ACTION A_PassEmsCmd:
// MQTT 명령 받기 (EMS 지령원이 있는 현장): GVL_IF.g_stEmsCmd를 번호를 확인하며 복사해 지령원 FB_SrcEms에 넘김 (GVL_IF 머리말의 읽는 규칙)
// 번호가 홀수 = 쓰는 중, 복사 전후 번호가 다름 = 복사 중에 바뀜 → 이번 스캔은 지난 복사본 그대로 (다음 스캔에 다시 시도)
nEmsSeq := GVL_IF.g_nCmdSeq;
// [결함 10 되돌림 2026-11-04: 코드로 막지 않고 운영 규칙으로 해결 — EMS는 command 토픽을 retain=false로 발행 (retained 명령은 재구독 때 새 메시지로 와서 실행됨).
//   되돌린 수정: IF (nEmsSeq AND 1) = 0 AND nEmsSeq <> 0 THEN (번호 0을 유효로 보지 않음) → 재시작 뒤 처음 온 정상 명령까지 번호 맞추기에만 쓰여 버려지는 부작용이 있었음]
IF (nEmsSeq AND 1) = 0 THEN
	stEmsCopy := GVL_IF.g_stEmsCmd;
	IF GVL_IF.g_nCmdSeq = nEmsSeq THEN
		GVL_SITE.g_fbSrcEms.i_stCmd		:= stEmsCopy;
		GVL_SITE.g_fbSrcEms.i_bValid	:= TRUE;
	END_IF
END_IF
GVL_SITE.g_fbSrcEms.i_astUnitCfg	:= GVL_SITE.UNIT_CFG;
GVL_SITE.g_fbSrcEms.i_astBmsCfg		:= GVL_SITE.BMS_CFG;
// 스탠다드 스케줄 모드: EMS PCS 지령을 그 PCS의 유닛에 넘김 (한 PCS에 유닛이 여럿이면 정격 비율로 나눔). 모드는 유닛별 값을 냄
// [16번 수정 2026-11-09: 관리자가 접속점 그룹 단위가 되어 모드 하나(g_fbCmStdSched1)가 모든 유닛 칸을 받음. 원래 g_fbCmStdSched1 ← PCS1, g_fbCmStdSched2 ← PCS2 그대로]
// 살아 있음 = EMS 지령원 유효 (지난 스캔). P 지령은 FB_SrcEms.i_bPEnable(기본 FALSE)과 따로라, 둘을 같이 켜지 않음
stEmsOut := GVL_SITE.g_fbSrcEms.Output;
FOR nCmU := 1 TO GVL_PARAM.UNIT_COUNT DO
	nCmPcs := GVL_SITE.UNIT_CFG[nCmU].nPcs;
	IF nCmPcs >= 1 AND nCmPcs <= GVL_PARAM.PCS_COUNT THEN
		fCmPcsRated := 0.0;
		FOR nCmK := 1 TO GVL_PARAM.UNIT_COUNT DO
			IF GVL_SITE.UNIT_CFG[nCmK].nPcs = nCmPcs AND F_RealOk(GVL_SITE.UNIT_CFG[nCmK].fPRated) THEN
				fCmPcsRated := fCmPcsRated + MAX(GVL_SITE.UNIT_CFG[nCmK].fPRated, 0.0);
			END_IF
		END_FOR
		GVL_SITE.g_fbCmStdSched1.i_astCmd[nCmU].bUse		:= TRUE;
		GVL_SITE.g_fbCmStdSched1.i_astCmd[nCmU].bAlive		:= stEmsOut.bValid;
		GVL_SITE.g_fbCmStdSched1.i_astCmd[nCmU].nPSeq		:= stEmsCopy.anPcsPSeq[nCmPcs];
		IF fCmPcsRated > 0.0 AND F_RealOk(GVL_SITE.UNIT_CFG[nCmU].fPRated) THEN
			GVL_SITE.g_fbCmStdSched1.i_astCmd[nCmU].fP	:= stEmsCopy.afPcsP[nCmPcs] * MAX(GVL_SITE.UNIT_CFG[nCmU].fPRated, 0.0) / fCmPcsRated;
		ELSE
			GVL_SITE.g_fbCmStdSched1.i_astCmd[nCmU].fP	:= 0.0;
		END_IF
		GVL_SITE.g_fbCmStdSched1.i_astCmd[nCmU].nStateSeq	:= stEmsCopy.astPcs[nCmPcs].nSeq;
		GVL_SITE.g_fbCmStdSched1.i_astCmd[nCmU].eState		:= stEmsCopy.astPcs[nCmPcs].eCmd;
	ELSE
		GVL_SITE.g_fbCmStdSched1.i_astCmd[nCmU].bUse		:= FALSE;	// PCS 번호 범위 밖 (설정 점검 오류)
	END_IF
END_FOR
END_ACTION

ACTION A_Report:
// UPS site: no installed PCS. Do not publish a Plaspo mapping for a UPS.
GVL_IF.g_nReportSeq:=GVL_IF.g_nReportSeq+1;
FOR _nReportPcs:=1 TO GVL_PARAM.PCS_COUNT DO
 GVL_IF.g_stReport.abPcsMapped[_nReportPcs]:=FALSE;
 GVL_IF.g_stReport.abPcsComm[_nReportPcs]:=FALSE;
END_FOR
fbRptBat[1](i_stState:=GVL_SITE.g_fbBms1.q_stState, i_stRaw:=GVL_SITE.g_fbBms1.q_stRaw, i_nDeviceIndex:=1);	// BAT 번호 1부터 [1부터 2026-11-10]
FOR _nReportBat:=1 TO GVL_PARAM.BMS_COUNT DO
 GVL_IF.g_stReport.abBatMapped[_nReportBat]:=TRUE;
 GVL_IF.g_stReport.abBatValid[_nReportBat]:=fbRptBat[_nReportBat].q_bValid;
 GVL_IF.g_stReport.astBat[_nReportBat]:=fbRptBat[_nReportBat].q_stBat;
 FOR _nReportRack:=1 TO GVL_PARAM.RACKS_PER_BMS DO
  GVL_IF.g_stReport.astRack[(_nReportBat-1)*GVL_PARAM.RACKS_PER_BMS+_nReportRack]:=fbRptBat[_nReportBat].q_astRack[_nReportRack];
 END_FOR
 FOR _nReportModule:=1 TO GVL_PARAM.RACKS_PER_BMS*GVL_PARAM.MODULES_PER_RACK DO
  GVL_IF.g_stReport.astModule[(_nReportBat-1)*GVL_PARAM.RACKS_PER_BMS*GVL_PARAM.MODULES_PER_RACK+_nReportModule]:=fbRptBat[_nReportBat].q_astModule[_nReportModule];
 END_FOR
END_FOR
fbRptUps[1](i_stState:=GVL_SITE.g_fbUps1.q_stState, i_nDeviceIndex:=1);
FOR _nReportUps:=1 TO GVL_PARAM.UPS_COUNT DO
 GVL_IF.g_stReport.abUpsMapped[_nReportUps]:=TRUE;
 GVL_IF.g_stReport.abUpsValid[_nReportUps]:=fbRptUps[_nReportUps].q_bValid;
 GVL_IF.g_stReport.astUps[_nReportUps]:=fbRptUps[_nReportUps].q_stUps;
 // 명세 SQ-01: 사고·고장 단계. Fault 확인 = EMS UPS 명령 10 (WR-SQ-01)
 fbUpsSafety[_nReportUps](i_stUps:=fbRptUps[_nReportUps].q_stUps, i_bUpsValid:=fbRptUps[_nReportUps].q_bValid,
  i_stBat:=fbRptBat[_nReportUps].q_stBat, i_bBatValid:=fbRptBat[_nReportUps].q_bValid, i_bAck:=fbUpsCommand[_nReportUps].q_bAck);
END_FOR
// IMD 보고 (인터페이스 22. IMD)
fbRptImd[1](i_stState:=GVL_SITE.g_fbImd1.q_stState, i_nDeviceIndex:=1);
FOR _nReportImd:=1 TO GVL_PARAM.IMD_COUNT DO
 GVL_IF.g_stReport.abImdMapped[_nReportImd]:=TRUE;
 GVL_IF.g_stReport.abImdValid[_nReportImd]:=fbRptImd[_nReportImd].q_bValid;
 GVL_IF.g_stReport.astImd[_nReportImd]:=fbRptImd[_nReportImd].q_stImd;
END_FOR
// 화재감지기 보고 (토픽 fire_detector, 인터페이스 20. OffGas 양식: b0 통신 이상, b1 알람, b2 고장)
// 1 = TS-60 연기 접점 (g_fbIo1 DI 1, 통신 = EtherCAT 단자 상태), 2 = ASD-57 (연기 또는 온도 알람). 고장(b2)은 알 수 없어 0
GVL_IF.g_stReport.abFireMapped[1]:=TRUE;
GVL_IF.g_stReport.astFire[1].DeviceIndex:=1;
GVL_IF.g_stReport.astFire[1].Status:=SEL(GVL_SITE.g_fbIo1.Comm, UDINT#1, SEL(GVL_SITE.g_fbIo1.M_GetBit(i_nPoint:=1), UDINT#0, UDINT#2));
GVL_IF.g_stReport.abFireMapped[2]:=TRUE;
GVL_IF.g_stReport.astFire[2].DeviceIndex:=2;
GVL_IF.g_stReport.astFire[2].Status:=SEL(GVL_SITE.g_fbAsd57.q_bValid, UDINT#1, SEL(GVL_SITE.g_fbAsd57.q_bSmokeAlarm OR GVL_SITE.g_fbAsd57.q_bTempAlarm, UDINT#0, UDINT#2));
// 온습도 보고 (인터페이스 07.Temperature Sensor). location 2 = BAT실 (잠정, 현장 위치 확인)
fbRptTemp[1](i_stState:=GVL_SITE.g_fbThd2.q_stState, i_nDeviceIndex:=1, i_nLocation:=2);
GVL_IF.g_stReport.abTempMapped[1]:=TRUE;
GVL_IF.g_stReport.astTemp[1]:=fbRptTemp[1].q_stTemp;
GVL_IF.g_nReportSeq:=GVL_IF.g_nReportSeq+1;
END_ACTION

END_PROGRAM

// ---- 10_Core/10_Snapshot/FB_Snapshot.TcPOU
FUNCTION_BLOCK FB_Snapshot		// 이번 스캔의 장비 상태를 한 번에 복사. 이후 단계는 이 사본만 읽는다
VAR_IN_OUT
	iq_aipPcs		: ARRAY[1..GVL_PARAM.PCS_COUNT] OF I_Pcs;
	iq_aipBms		: ARRAY[1..GVL_PARAM.BMS_COUNT] OF I_Bms;
	iq_aipMeter		: ARRAY[1..GVL_PARAM.METER_COUNT] OF I_Meter;
END_VAR
VAR_IN_OUT CONSTANT
	iq_astUnitCfg	: ARRAY[1..GVL_PARAM.UNIT_COUNT] OF ST_UnitCfg;
END_VAR
VAR_OUTPUT
	q_astUnit		: ARRAY[1..GVL_PARAM.UNIT_COUNT] OF ST_UnitState;
	q_astBms		: ARRAY[1..GVL_PARAM.BMS_COUNT] OF ST_BatState;
	q_astMeter		: ARRAY[1..GVL_PARAM.METER_COUNT] OF ST_MeterState;
END_VAR
VAR_TEMP
	i				: UINT;
	nPcs			: UINT;
	stNoUnit		: ST_UnitState;		// 빈 칸: 통신 없음, 상태 Unknown
	stNoBms			: ST_BatState;
	stNoMeter		: ST_MeterState;
	k				: UINT;		// [결함 9 수정 2026-11-03: 추가]
END_VAR

// 유닛: 구성표의 PCS 번호·PCS 안 번호로 찾음
FOR i := 1 TO GVL_PARAM.UNIT_COUNT DO
	nPcs := iq_astUnitCfg[i].nPcs;
	IF nPcs >= 1 AND nPcs <= GVL_PARAM.PCS_COUNT AND_THEN iq_aipPcs[nPcs] <> 0 THEN
		q_astUnit[i] := iq_aipPcs[nPcs].M_GetUnitState(iq_astUnitCfg[i].nSub);
		q_astUnit[i].stP := M_FixVal(q_astUnit[i].stP);	// [결함 9 수정 2026-11-03: NaN·무한대 → 0·무효]
		q_astUnit[i].stQ := M_FixVal(q_astUnit[i].stQ);
	ELSE
		q_astUnit[i] := stNoUnit;
	END_IF
END_FOR

FOR i := 1 TO GVL_PARAM.BMS_COUNT DO
	IF iq_aipBms[i] <> 0 THEN
		q_astBms[i] := iq_aipBms[i].BatState;
		q_astBms[i].stSoc := M_FixVal(q_astBms[i].stSoc);	// [결함 9 수정 2026-11-03: NaN·무한대 → 0·무효, 한도는 0]
		q_astBms[i].stSoh := M_FixVal(q_astBms[i].stSoh);
		IF NOT F_CmdOk(q_astBms[i].fPChgMax, 0.0) THEN q_astBms[i].fPChgMax := 0.0; END_IF
		IF NOT F_CmdOk(q_astBms[i].fPDisMax, 0.0) THEN q_astBms[i].fPDisMax := 0.0; END_IF
	ELSE
		q_astBms[i] := stNoBms;
	END_IF
END_FOR

FOR i := 1 TO GVL_PARAM.METER_COUNT DO
	IF iq_aipMeter[i] <> 0 THEN
		q_astMeter[i] := iq_aipMeter[i].MeterState;
		q_astMeter[i].stP := M_FixVal(q_astMeter[i].stP);	// [결함 9 수정 2026-11-03: NaN·무한대 → 0·무효]
		q_astMeter[i].stQ := M_FixVal(q_astMeter[i].stQ);
		q_astMeter[i].stV := M_FixVal(q_astMeter[i].stV);
		FOR k := 1 TO 3 DO
			q_astMeter[i].astV[k] := M_FixVal(q_astMeter[i].astV[k]);
		END_FOR
		q_astMeter[i].stF := M_FixVal(q_astMeter[i].stF);
	ELSE
		q_astMeter[i] := stNoMeter;
	END_IF
END_FOR

METHOD PRIVATE M_FixVal : ST_Val		// 장비 값이 NaN·무한대면 0·무효로 (뒤 계산·비교에 퍼지지 않게). [결함 9 수정 2026-11-03: 추가]
VAR_INPUT
	i_stVal	: ST_Val;
END_VAR
M_FixVal := i_stVal;
IF NOT F_CmdOk(i_stVal.fValue, 0.0) THEN
	M_FixVal.fValue	:= 0.0;
	M_FixVal.bValid	:= FALSE;
END_IF
END_METHOD

END_FUNCTION_BLOCK

// ---- 10_Core/40_Arbitration/F_CmdOk.TcPOU
FUNCTION F_CmdOk : BOOL		// 지령값이 쓸 만한가: NaN·무한대가 아니고, 한도가 있으면 |값| ≤ 한도
VAR_INPUT
	i_fValue	: REAL;
	i_fLimit	: REAL;			// 0 이하 = 한도 검사 안 함
END_VAR

// NaN·무한대는 비트로 먼저 거름 (NaN을 크기 비교하면 PLC가 멈춤). 크기 비교는 보통 숫자일 때만
// [2026-11-05 머지: main의 F_IsFinite 방식 + 1.0E30 상한은 원래 코드대로 남김. 통합시험 결함 9 수정(비트 검사·dwBits)은 이 방식으로 합침]
F_CmdOk := F_IsFinite(i_fValue) AND_THEN ABS(i_fValue) < 1.0E30;
IF F_CmdOk AND i_fLimit > 0 THEN
	F_CmdOk := ABS(i_fValue) <= i_fLimit;
END_IF

END_FUNCTION

// ---- 10_Core/10_Snapshot/FB_Measure.TcPOU
FUNCTION_BLOCK FB_Measure		// 계측점 계산 + 제어 그룹마다 접속점 값·가상신호
VAR_INPUT
	i_bTestMode		: BOOL;			// 시험 모드에서만 가상신호를 씀 (GVL_SITE.TEST_MODE)
END_VAR
VAR_IN_OUT CONSTANT
	iq_astMeter		: ARRAY[1..GVL_PARAM.METER_COUNT] OF ST_MeterState;
	iq_astPointCfg	: ARRAY[1..GVL_PARAM.POINT_COUNT] OF ST_PointCfg;
	iq_astGroupCfg	: ARRAY[1..GVL_PARAM.GROUP_COUNT] OF ST_GroupCfg;
	iq_astVirtual	: ARRAY[1..GVL_PARAM.GROUP_COUNT] OF ST_VirtualSet;
END_VAR
VAR_OUTPUT
	q_astPoint		: ARRAY[1..GVL_PARAM.POINT_COUNT] OF ST_MeterState;	// 계측점 (실측, 가상신호 적용 전)
	q_astPcc		: ARRAY[1..GVL_PARAM.GROUP_COUNT] OF ST_PccMeas;		// 그룹 접속점 (가상신호 적용 후)
END_VAR
VAR_TEMP
	nPointNo				: UINT;
	nTermNo				: UINT;
	g				: UINT;
	k				: UINT;
	nMeterNo				: UINT;
	bFirst			: BOOL;		// 아직 묶인 계측기를 못 만남
	bComm			: BOOL;
	bPValid			: BOOL;
	bQValid			: BOOL;
	stPoint			: ST_MeterState;
	stNone			: ST_MeterState;	// 빈 값: 통신 없음, 값 무효
END_VAR

(* 1) 계측점: 계측기 P·Q를 부호와 함께 더함. 전압·주파수는 첫 계측기 값 *)
FOR nPointNo := 1 TO GVL_PARAM.POINT_COUNT DO
	stPoint	:= stNone;
	bFirst	:= TRUE;
	bComm	:= TRUE;
	bPValid	:= TRUE;
	bQValid	:= TRUE;
	FOR nTermNo := 1 TO GVL_PARAM.POINT_TERM_MAX DO
		nMeterNo := iq_astPointCfg[nPointNo].astTerm[nTermNo].nMeter;
		IF nMeterNo > GVL_PARAM.METER_COUNT THEN
			bComm := FALSE;		// 설정 오류: 없는 계측기
		ELSIF nMeterNo >= 1 THEN
			IF bFirst THEN
				stPoint.stV	:= iq_astMeter[nMeterNo].stV;
				stPoint.astV	:= iq_astMeter[nMeterNo].astV;
				stPoint.stF	:= iq_astMeter[nMeterNo].stF;
				bFirst		:= FALSE;
			END_IF
			bComm			:= bComm AND iq_astMeter[nMeterNo].bComm;
			bPValid			:= bPValid AND iq_astMeter[nMeterNo].stP.bValid;
			bQValid			:= bQValid AND iq_astMeter[nMeterNo].stQ.bValid;
			stPoint.stP.fValue	:= stPoint.stP.fValue + iq_astPointCfg[nPointNo].astTerm[nTermNo].fSign * iq_astMeter[nMeterNo].stP.fValue;
			stPoint.stQ.fValue	:= stPoint.stQ.fValue + iq_astPointCfg[nPointNo].astTerm[nTermNo].fSign * iq_astMeter[nMeterNo].stQ.fValue;
		END_IF
	END_FOR
	// 묶인 계측기가 없거나 하나라도 끊기면 무효
	stPoint.bComm		:= bComm AND NOT bFirst;
	stPoint.stP.bValid	:= stPoint.bComm AND bPValid;
	stPoint.stQ.bValid	:= stPoint.bComm AND bQValid;
	q_astPoint[nPointNo]	:= stPoint;
END_FOR

(* 2) 그룹 접속점 + 가상신호 *)
FOR g := 1 TO GVL_PARAM.GROUP_COUNT DO
	nPointNo := iq_astGroupCfg[g].nPccPoint;
	q_astPcc[g].bNoPoint := nPointNo = 0;	// [결함 7 수정 2026-11-03: 추가. 접속점 무효 보호가 '없음'을 무효로 보지 않게]
	IF nPointNo >= 1 AND nPointNo <= GVL_PARAM.POINT_COUNT THEN
		q_astPcc[g].stMeas := q_astPoint[nPointNo];
	ELSE
		q_astPcc[g].stMeas := stNone;
	END_IF

	// 가상 전압: 평균·상전압 모두 같은 값
	IF i_bTestMode AND iq_astVirtual[g].bVEna THEN
		q_astPcc[g].stMeas.stV.fValue	:= iq_astVirtual[g].fV;
		q_astPcc[g].stMeas.stV.bValid	:= TRUE;
		FOR k := 1 TO 3 DO
			q_astPcc[g].stMeas.astV[k].fValue	:= iq_astVirtual[g].fV;
			q_astPcc[g].stMeas.astV[k].bValid	:= TRUE;
		END_FOR
	END_IF

	// 가상 유효전력
	IF i_bTestMode AND iq_astVirtual[g].bPEna THEN
		q_astPcc[g].stMeas.stP.fValue	:= iq_astVirtual[g].fP;
		q_astPcc[g].stMeas.stP.bValid	:= TRUE;
	END_IF
END_FOR

END_FUNCTION_BLOCK

// ---- 10_Core/20_Protection/FB_Protection.TcPOU
FUNCTION_BLOCK FB_Protection		// 등록된 보호 칸마다 대상마다: 조건 모듈 판단 → 같은 칸 대응 모듈 → 유닛·BMS마다 요청 합치기 (센 조치·낮은 상한, 건 모듈 ID). 요청만, 장비에 직접 명령하지 않음
// 지연 없음: 통신 에러·고장은 장비 쪽(드라이버)이 판정해 올림. 현장 접점·아날로그의 떨림 방지는 조건 모듈 설정에
// 보호는 조건이 있는 동안만 걸림 (래치 없음). 다시 돌지 않아야 하면 정지나 Manual 전환을 씀
VAR_IN_OUT CONSTANT
	iq_astUnit		: ARRAY[1..GVL_PARAM.UNIT_COUNT] OF ST_UnitState;
	iq_astBms		: ARRAY[1..GVL_PARAM.BMS_COUNT] OF ST_BatState;
	iq_astPcc		: ARRAY[1..GVL_PARAM.GROUP_COUNT] OF ST_PccMeas;
	iq_astUnitCfg	: ARRAY[1..GVL_PARAM.UNIT_COUNT] OF ST_UnitCfg;
	iq_astBmsCfg	: ARRAY[1..GVL_PARAM.BMS_COUNT] OF ST_BmsCfg;
	iq_astRuleCfg	: ARRAY[1..GVL_PARAM.RULE_COUNT] OF ST_RuleCfg;
	iq_abUnitInstalled	: ARRAY[1..GVL_PARAM.UNIT_COUNT] OF BOOL;	// 미설치(칸 비어 있음)는 모듈에 bInstalled = FALSE로 넘김 (FB_ModuleList)
	iq_abBmsInstalled	: ARRAY[1..GVL_PARAM.BMS_COUNT] OF BOOL;
	iq_aeOpMode		: ARRAY[1..GVL_PARAM.UNIT_COUNT] OF E_OpMode;		// 실제 운전 모드 (대응이 그 모드 유닛에 조치를 걸지 봄)
END_VAR
VAR_IN_OUT
	iq_aipRule		: ARRAY[1..GVL_PARAM.RULE_COUNT] OF I_ProtectionRule;	// 조건 모듈
	iq_aipResp		: ARRAY[1..GVL_PARAM.RULE_COUNT] OF I_ProtResponse;	// 대응 모듈 (같은 칸). 비우면 조치 없음 (알람만)
END_VAR
VAR_OUTPUT
	q_astUnitProt	: ARRAY[1..GVL_PARAM.UNIT_COUNT] OF ST_UnitProt;		// 유닛별 가장 센 PCS 조치·가장 낮은 P·Q 상한·Manual 전환
	q_astBmsProt	: ARRAY[1..GVL_PARAM.BMS_COUNT] OF ST_BmsProt;		// BMS별 가장 센 배터리 조치
	q_aabRule		: ARRAY[1..GVL_PARAM.RULE_COUNT, 1..GVL_PARAM.PROT_TARGET_MAX] OF BOOL;	// 보호 발생 [규칙 칸, 대상 번호] (온라인 확인·로그용). Site는 대상 1
END_VAR
VAR
	_aatonActive	: ARRAY[1..GVL_PARAM.RULE_COUNT, 1..GVL_PARAM.PROT_TARGET_MAX] OF TON;	// 조건이 이어진 시간 (대응에 넘김)
	_stView			: ST_ProtView;		// 마지막으로 조건 모듈에 넘긴 정보 (온라인 확인용)
	_stReq			: ST_ProtReq;		// 마지막 대응 요청 (온라인 확인용)
	_stNoReq		: ST_ProtReq;		// 요청 없음 (비우기용. 처음 한 번 P·Q 상한을 100으로)
	_bInit			: BOOL;
END_VAR
VAR_TEMP
	i				: UINT;		// 규칙 칸
	t				: UINT;		// 대상 번호
	nTargetCount	: UINT;		// 이 규칙 범위의 대상 수
	bInRange		: BOOL;		// 이 대상을 보는가
	bCond			: BOOL;
	nModule			: UINT;
	stNoUnit		: ST_UnitProt;
	stNoBms			: ST_BmsProt;
	stNoView		: ST_ProtView;
END_VAR

(* 0) 이번 스캔 결과 비우기 *)
IF NOT _bInit THEN
	FOR i := 1 TO GVL_PARAM.UNIT_COUNT DO
		_stNoReq.afPPct[i] := 100.0;
		_stNoReq.afQPct[i] := 100.0;
	END_FOR
	_bInit := TRUE;
END_IF
FOR i := 1 TO GVL_PARAM.UNIT_COUNT DO
	q_astUnitProt[i] := stNoUnit;
END_FOR
FOR i := 1 TO GVL_PARAM.BMS_COUNT DO
	q_astBmsProt[i] := stNoBms;
END_FOR
(* 1) 보호 규칙 칸마다, 범위 안 대상마다: 조건 모듈 → 대응 → 합치기
   대상 번호(nTarget) 0 = 범위 안 대상 전부를 하나씩 (유닛 범위면 유닛 1..UNIT_COUNT). Site는 대상 1 하나 *)
FOR i := 1 TO GVL_PARAM.RULE_COUNT DO
	CASE iq_astRuleCfg[i].eScope OF
		E_ProtScope.Unit:		nTargetCount := GVL_PARAM.UNIT_COUNT;
		E_ProtScope.Bms:		nTargetCount := GVL_PARAM.BMS_COUNT;
		E_ProtScope.BatGroup:	nTargetCount := GVL_PARAM.BAT_COUNT;
		E_ProtScope.Group:		nTargetCount := GVL_PARAM.GROUP_COUNT;
	ELSE
		nTargetCount := 1;		// Site
	END_CASE
	nModule := 0;
	IF iq_aipRule[i] <> 0 THEN
		nModule := iq_aipRule[i].ModuleId;
	END_IF
	FOR t := 1 TO GVL_PARAM.PROT_TARGET_MAX DO
		bInRange := iq_aipRule[i] <> 0 AND t <= nTargetCount
			AND (iq_astRuleCfg[i].nTarget = 0 OR iq_astRuleCfg[i].nTarget = t OR iq_astRuleCfg[i].eScope = E_ProtScope.Site);
		bCond := FALSE;
		IF bInRange THEN
			// 조건 모듈에 넘길 정보: 범위·대상 번호·임계값과 그 대상의 상태
			_stView				:= stNoView;
			_stView.eScope		:= iq_astRuleCfg[i].eScope;
			_stView.nTarget		:= t;
			_stView.fThreshold	:= iq_astRuleCfg[i].fThreshold;
			_stView.bInstalled	:= TRUE;
			CASE iq_astRuleCfg[i].eScope OF
				E_ProtScope.Unit:
					_stView.bInstalled	:= iq_abUnitInstalled[t];
					_stView.stUnit		:= iq_astUnit[t];
					_stView.eOpMode		:= iq_aeOpMode[t];
					_stView.nGroup		:= iq_astUnitCfg[t].nGroup;
					_stView.nBatGroup	:= iq_astUnitCfg[t].nBatGroup;
				E_ProtScope.Bms:
					_stView.bInstalled	:= iq_abBmsInstalled[t];
					_stView.stBms		:= iq_astBms[t];
					_stView.nBatGroup	:= iq_astBmsCfg[t].nBatGroup;
				E_ProtScope.BatGroup:
					_stView.nBatGroup	:= t;
				E_ProtScope.Group:
					_stView.stPcc		:= iq_astPcc[t];
					_stView.nGroup		:= t;
			END_CASE
			// 등록 bAuto·bManual 중 하나라도 켜져 있어야 감지 (둘 다 끄면 이 보호를 안 씀)
			bCond := (iq_astRuleCfg[i].stProt.bAuto OR iq_astRuleCfg[i].stProt.bManual) AND iq_aipRule[i].M_Evaluate(_stView);
		END_IF
		q_aabRule[i, t] := bCond;
		_aatonActive[i, t](IN := bCond, PT := T#24D);
		// 대응: 매 스캔 부름 (조건이 없을 때도: 단계 대응이 풀린 뒤 상태를 정리할 수 있게). 대응 칸이 비면 조치 없음 (알람만)
		IF bInRange AND iq_aipResp[i] <> 0 THEN
			_stReq := _stNoReq;
			iq_aipResp[i].M_Respond(i_bActive := bCond, i_tActive := _aatonActive[i, t].ET, i_nTarget := t, i_stRule := iq_astRuleCfg[i],
				iq_astUnit := iq_astUnit, iq_astBms := iq_astBms, iq_astUnitCfg := iq_astUnitCfg, iq_astBmsCfg := iq_astBmsCfg,
				iq_aeOpMode := iq_aeOpMode, iq_stReq := _stReq);
			M_Merge(nModule);
		END_IF
	END_FOR
END_FOR

METHOD PRIVATE M_Merge		// 대응 요청(_stReq)을 장비마다 합침: PCS·배터리는 센 쪽, P·Q 상한은 낮은 쪽, Manual 전환은 하나라도. 건 모듈 = 조건 모듈 ID
VAR_INPUT
	i_nModule	: UINT;
END_VAR
VAR
	u			: UINT;
	m			: UINT;
END_VAR
FOR u := 1 TO GVL_PARAM.UNIT_COUNT DO
	IF F_PcsRank(_stReq.aePcs[u]) > F_PcsRank(q_astUnitProt[u].ePcsAction) THEN
		q_astUnitProt[u].ePcsAction	:= _stReq.aePcs[u];
		q_astUnitProt[u].nModule	:= i_nModule;
	END_IF
	IF _stReq.abToManual[u] AND NOT q_astUnitProt[u].bModeManualReq THEN
		q_astUnitProt[u].bModeManualReq	:= TRUE;
		q_astUnitProt[u].nModeModule	:= i_nModule;
	END_IF
	IF _stReq.afPPct[u] < q_astUnitProt[u].fPPct THEN
		q_astUnitProt[u].fPPct		:= _stReq.afPPct[u];
		q_astUnitProt[u].nPModule	:= i_nModule;
	END_IF
	IF _stReq.afQPct[u] < q_astUnitProt[u].fQPct THEN
		q_astUnitProt[u].fQPct		:= _stReq.afQPct[u];
		q_astUnitProt[u].nQModule	:= i_nModule;
	END_IF
END_FOR
FOR m := 1 TO GVL_PARAM.BMS_COUNT DO
	IF F_BatRank(_stReq.aeBat[m]) > F_BatRank(q_astBmsProt[m].eBatAction) THEN
		q_astBmsProt[m].eBatAction	:= _stReq.aeBat[m];
		q_astBmsProt[m].nModule		:= i_nModule;
	END_IF
END_FOR
END_METHOD

END_FUNCTION_BLOCK

// ---- 10_Core/20_Protection/F_PcsRank.TcPOU
FUNCTION F_PcsRank : INT		// 조치 세기: None 0 < Standby 1 < Stop 2 < EStop 3
VAR_INPUT
	i_eAction	: E_PcsAction;
END_VAR

CASE i_eAction OF
	E_PcsAction.Standby:	F_PcsRank := 1;
	E_PcsAction.Stop:		F_PcsRank := 2;
	E_PcsAction.EStop:		F_PcsRank := 3;
ELSE
	F_PcsRank := 0;
END_CASE

END_FUNCTION

// ---- 10_Core/20_Protection/F_BatRank.TcPOU
FUNCTION F_BatRank : INT		// 조치 세기: None 0 < Stop 1 < EStop 2
VAR_INPUT
	i_eAction	: E_BatAction;
END_VAR

CASE i_eAction OF
	E_BatAction.Stop:	F_BatRank := 1;
	E_BatAction.EStop:	F_BatRank := 2;
ELSE
	F_BatRank := 0;
END_CASE

END_FUNCTION

// ---- 10_Core/20_Protection/FB_BatGroup.TcPOU
FUNCTION_BLOCK FB_BatGroup		// BMS마다 쓸 수 있는지 판단, 배터리 그룹(DC 버스)마다 쓸 수 있는 BMS만 모음 (한도·SOC·투입 완료)
VAR_IN_OUT CONSTANT
	iq_astBms		: ARRAY[1..GVL_PARAM.BMS_COUNT] OF ST_BatState;
	iq_astBmsCfg	: ARRAY[1..GVL_PARAM.BMS_COUNT] OF ST_BmsCfg;
	iq_astBmsProt	: ARRAY[1..GVL_PARAM.BMS_COUNT] OF ST_BmsProt;
	iq_abBmsInstalled	: ARRAY[1..GVL_PARAM.BMS_COUNT] OF BOOL;	// FB_ModuleList. 미설치 BMS는 배터리 그룹에서 뺌
END_VAR
VAR_OUTPUT
	q_astBmsAvail	: ARRAY[1..GVL_PARAM.BMS_COUNT] OF ST_BmsAvail;
	q_astBatGroup	: ARRAY[1..GVL_PARAM.BAT_COUNT] OF ST_BatGroupState;
END_VAR
VAR_TEMP
	m				: UINT;
	g				: UINT;
	fCapWeight				: REAL;		// 무게 = 용량 (설정 안 했으면 1)
	fSocW			: REAL;
	fWSum			: REAL;
	nClosed			: UINT;		// 쓸 수 있는 BMS 중 투입된 수
	fChgClosed		: REAL;		// 투입된 BMS 한도 합 (투입된 BMS가 있으면 이것만 씀: 열린 BMS 한도로 과부하 안 되게)
	fDisClosed		: REAL;
	stBmsAvail			: ST_BmsAvail;
	stBmsAvailNone		: ST_BmsAvail;
	stGrp				: ST_BatGroupState;
	stNone			: ST_BatGroupState;
END_VAR

(* 1) BMS마다 쓸 수 있는지 *)
FOR m := 1 TO GVL_PARAM.BMS_COUNT DO
	stBmsAvail			:= stBmsAvailNone;
	stBmsAvail.bNotInstalled	:= NOT iq_abBmsInstalled[m];
	stBmsAvail.bNoComm	:= iq_abBmsInstalled[m] AND NOT iq_astBms[m].bComm;
	stBmsAvail.bFault		:= iq_astBms[m].bComm AND iq_astBms[m].bFault;
	stBmsAvail.bSysStop	:= iq_astBms[m].bComm AND iq_astBms[m].bSysStop;
	stBmsAvail.bProt		:= iq_astBmsProt[m].eBatAction <> E_BatAction.None;
	stBmsAvail.bUsable	:= NOT (stBmsAvail.bNotInstalled OR stBmsAvail.bNoComm OR stBmsAvail.bFault OR stBmsAvail.bSysStop OR stBmsAvail.bProt);
	q_astBmsAvail[m] := stBmsAvail;
END_FOR

(* 2) 배터리 그룹마다 쓸 수 있는 BMS만 합침 *)
FOR g := 1 TO GVL_PARAM.BAT_COUNT DO
	stGrp		:= stNone;
	fSocW	:= 0;
	fWSum	:= 0;
	nClosed	:= 0;
	fChgClosed	:= 0;
	fDisClosed	:= 0;
	FOR m := 1 TO GVL_PARAM.BMS_COUNT DO
		IF iq_astBmsCfg[m].nBatGroup = g AND iq_abBmsInstalled[m] THEN
			stGrp.nBms := stGrp.nBms + 1;
			IF q_astBmsAvail[m].bUsable THEN
				stGrp.nBmsUsable	:= stGrp.nBmsUsable + 1;
				IF iq_astBms[m].bContactorClosed THEN
					nClosed		:= nClosed + 1;
					fChgClosed	:= fChgClosed + iq_astBms[m].fPChgMax;
					fDisClosed	:= fDisClosed + iq_astBms[m].fPDisMax;
				END_IF
				stGrp.fPChgMax		:= stGrp.fPChgMax + iq_astBms[m].fPChgMax;
				stGrp.fPDisMax		:= stGrp.fPDisMax + iq_astBms[m].fPDisMax;
				IF iq_astBms[m].stSoc.bValid THEN
					fCapWeight := SEL(iq_astBmsCfg[m].fCapacity > 0, 1.0, iq_astBmsCfg[m].fCapacity);
					IF fWSum = 0 OR iq_astBms[m].stSoc.fValue < stGrp.stSocMin.fValue THEN stGrp.stSocMin.fValue := iq_astBms[m].stSoc.fValue; END_IF
					IF fWSum = 0 OR iq_astBms[m].stSoc.fValue > stGrp.stSocMax.fValue THEN stGrp.stSocMax.fValue := iq_astBms[m].stSoc.fValue; END_IF
					fSocW	:= fSocW + iq_astBms[m].stSoc.fValue * fCapWeight;
					fWSum	:= fWSum + fCapWeight;
					stGrp.fCapacity	:= stGrp.fCapacity + MAX(iq_astBmsCfg[m].fCapacity, 0.0);	// SOC 평균에 들어간 BMS만 (용량 × SOC = 에너지가 맞게)
				END_IF
			END_IF
		END_IF
	END_FOR
	IF fWSum > 0 THEN
		stGrp.stSoc.fValue		:= fSocW / fWSum;
		stGrp.stSoc.bValid		:= TRUE;
		stGrp.stSocMin.bValid	:= TRUE;
		stGrp.stSocMax.bValid	:= TRUE;
		stGrp.fSocWeight		:= fWSum;
	END_IF
	// 한도: 투입된 BMS가 있으면 그 BMS 것만 (열린 BMS는 전류를 못 받음). 하나도 없으면(기동 전) 쓸 수 있는 BMS 전부 (화면·판단용, 그대로)
	IF nClosed > 0 THEN
		stGrp.fPChgMax := fChgClosed;
		stGrp.fPDisMax := fDisClosed;
	END_IF
	stGrp.bUsable := stGrp.nBmsUsable > 0;
	stGrp.bReady := stGrp.nBmsUsable > 0 AND nClosed = stGrp.nBmsUsable;
	q_astBatGroup[g] := stGrp;
END_FOR

END_FUNCTION_BLOCK

// ---- 10_Core/20_Protection/FB_UnitAvail.TcPOU
FUNCTION_BLOCK FB_UnitAvail		// 유닛마다 쓸 수 있는 상태인지와 그 이유 (통신·고장·로컬·배터리·보호)
VAR_IN_OUT CONSTANT
	iq_astUnit		: ARRAY[1..GVL_PARAM.UNIT_COUNT] OF ST_UnitState;
	iq_astUnitCfg	: ARRAY[1..GVL_PARAM.UNIT_COUNT] OF ST_UnitCfg;
	iq_astUnitProt	: ARRAY[1..GVL_PARAM.UNIT_COUNT] OF ST_UnitProt;
	iq_astBatGroup	: ARRAY[1..GVL_PARAM.BAT_COUNT] OF ST_BatGroupState;
	iq_abUnitInstalled	: ARRAY[1..GVL_PARAM.UNIT_COUNT] OF BOOL;	// FB_ModuleList. 미설치 유닛은 가용 아님 (이유 bNotInstalled만)
END_VAR
VAR_OUTPUT
	q_astAvail		: ARRAY[1..GVL_PARAM.UNIT_COUNT] OF ST_UnitAvail;
END_VAR
VAR_TEMP
	u				: UINT;
	b				: UINT;
	stUnitAvail			: ST_UnitAvail;
	stNone			: ST_UnitAvail;
END_VAR

FOR u := 1 TO GVL_PARAM.UNIT_COUNT DO
	stUnitAvail := stNone;

	// PCS (미설치면 통신·고장 판단을 안 함)
	stUnitAvail.bNotInstalled	:= NOT iq_abUnitInstalled[u];
	stUnitAvail.bNoPcsComm	:= iq_abUnitInstalled[u] AND NOT iq_astUnit[u].bComm;
	stUnitAvail.bPcsFault	:= iq_astUnit[u].bComm AND iq_astUnit[u].bFault;
	stUnitAvail.bPcsLocal	:= F_IsLocal(iq_astUnit[u]);
	stUnitAvail.bProt		:= iq_astUnitProt[u].ePcsAction <> E_PcsAction.None;

	// 연결 배터리 그룹 (0 = 배터리 없는 유닛)
	b := iq_astUnitCfg[u].nBatGroup;
	IF b > GVL_PARAM.BAT_COUNT THEN
		stUnitAvail.bNoBat := TRUE;		// 설정 오류
	ELSIF b >= 1 THEN
		stUnitAvail.bNoBat := NOT iq_astBatGroup[b].bUsable;
	END_IF

	stUnitAvail.bAvail := NOT (stUnitAvail.bNotInstalled OR stUnitAvail.bNoPcsComm OR stUnitAvail.bPcsFault OR stUnitAvail.bPcsLocal OR stUnitAvail.bNoBat OR stUnitAvail.bProt);
	q_astAvail[u] := stUnitAvail;
END_FOR

END_FUNCTION_BLOCK

// ---- 10_Core/02_Util/F_IsLocal.TcPOU
FUNCTION F_IsLocal : BOOL		// PCS가 로컬(PMS 제어 안 받음)인가. 통신이 끊긴 건 로컬로 보지 않음
VAR_INPUT
	i_stUnit	: ST_UnitState;
END_VAR

F_IsLocal := i_stUnit.bComm AND NOT i_stUnit.bCtrlReady;

END_FUNCTION

// ---- 10_Core/20_Protection/FB_EquipmentLimits.TcPOU
FUNCTION_BLOCK FB_EquipmentLimits	// 설비 한도: 유닛(정격 × Derate ∩ 유닛 제한 모듈), 배터리 버스(BMS 한도 ∩ 버스 제한 모듈), 그룹 설비 범위. 스캔당 한 번
// 성형(그룹 설비 범위)과 분배(유닛·버스 한도)가 이 결과를 같이 씀: 같은 한도를 두 곳에서 따로 계산하지 않음
// 모듈은 범위를 좁히기만 함 (넓힐 수 없음). 0은 항상 범위 안 (모듈이 출력을 강제하지 못함)
// 유닛 제한은 유닛의 실제 운전 모드에 맞는 등록(bAuto·bManual)만, 버스 제한은 그 버스에 대상 모드 유닛이 하나라도 있으면 버스 전체에 건다
VAR_IN_OUT CONSTANT
	iq_astUnitCfg	: ARRAY[1..GVL_PARAM.UNIT_COUNT] OF ST_UnitCfg;
	iq_astUnit	: ARRAY[1..GVL_PARAM.UNIT_COUNT] OF ST_UnitState;
	iq_astAvail	: ARRAY[1..GVL_PARAM.UNIT_COUNT] OF ST_UnitAvail;
	iq_astUnitProt	: ARRAY[1..GVL_PARAM.UNIT_COUNT] OF ST_UnitProt;	// 보호 Derate
	iq_aeOpMode	: ARRAY[1..GVL_PARAM.UNIT_COUNT] OF E_OpMode;	// 실제 운전 모드
	iq_astBatGroup	: ARRAY[1..GVL_PARAM.BAT_COUNT] OF ST_BatGroupState;
	iq_astUnitRuleReg	: ARRAY[1..GVL_PARAM.UNIT_RULE_COUNT] OF ST_RuleTargetReg;
	iq_astBatRuleReg	: ARRAY[1..GVL_PARAM.BAT_RULE_COUNT] OF ST_RuleTargetReg;
END_VAR
VAR_IN_OUT
	iq_aipUnitRule	: ARRAY[1..GVL_PARAM.UNIT_RULE_COUNT] OF I_UnitLimitRule;
	iq_aipBatRule	: ARRAY[1..GVL_PARAM.BAT_RULE_COUNT] OF I_BatLimitRule;
END_VAR
VAR_OUTPUT
	q_astUnitEnv	: ARRAY[1..GVL_PARAM.UNIT_COUNT] OF ST_UnitEnvelope;	// 유닛 한도 (분배)
	q_astBatEnv	: ARRAY[1..GVL_PARAM.BAT_COUNT] OF ST_BatEnvelope;	// 버스 한도 (분배)
	q_astGroupEnv	: ARRAY[1..GVL_PARAM.GROUP_COUNT] OF ST_GroupEnvelope;	// 그룹 설비 범위 (성형)
END_VAR
VAR
	(* 반복 변수·임시값: 본문과 액션(A_)이 함께 씀. 액션이 본문의 VAR_TEMP를 못 볼 수 있어 VAR에 둠 *)
	_u	: UINT;
	_b	: UINT;
	_g	: UINT;
	_i	: UINT;
	_bManual	: BOOL;
	_fRatio	: REAL;
	_fSP	: REAL;		// kW, 보호 P 상한 (정격 × P%). 피상전력 상한 계산용
	_fSQ	: REAL;		// kvar, 보호 Q 상한 (정격 × Q%). 피상전력 상한 계산용
	_stUnitView	: ST_UnitLimitView;
	_stBatView	: ST_BatLimitView;
	_stLimOut	: ST_LimitOut;
	_stBatOut	: ST_BatLimitOut;
	_stEnv	: ST_UnitEnvelope;
	_stEnvNone	: ST_UnitEnvelope;
	_stBatEnv	: ST_BatEnvelope;
	_stBatNone	: ST_BatEnvelope;
	_stGrp	: ST_GroupEnvelope;
	_stGrpNone	: ST_GroupEnvelope;
	_stNew	: ST_Range;
	_stNoVal	: ST_Val;
	_anAuto	: ARRAY[1..GVL_PARAM.BAT_COUNT] OF UINT;	// 버스의 Auto 유닛 수
	_anManual	: ARRAY[1..GVL_PARAM.BAT_COUNT] OF UINT;	// 버스의 Manual 유닛 수
	_afBusOut	: ARRAY[1..GVL_PARAM.BAT_COUNT] OF REAL;	// 버스 유닛 실측 P 합
	_afBusMax	: ARRAY[1..GVL_PARAM.BAT_COUNT] OF REAL;	// 이 그룹 가용 유닛 P 상한 합 (버스별)
	_afBusMin	: ARRAY[1..GVL_PARAM.BAT_COUNT] OF REAL;
	_abBusIn	: ARRAY[1..GVL_PARAM.BAT_COUNT] OF BOOL;	// 이 그룹 가용 유닛이 쓰는 버스
END_VAR

A_CountBusUnit();		// 버스마다 운전 모드별 유닛 수, 출력 합
A_CalcBusLimit();		// 버스 한도: BMS 한도 합 ∩ 버스 제한 모듈
A_CalcUnitLimit();		// 유닛 한도: 정격 × Derate ∩ 유닛 제한 모듈
A_CalcGroupRange();		// 그룹 설비 범위 (가용 유닛)

ACTION A_CountBusUnit:
(* 1) 버스마다 운전 모드별 유닛 수, 출력 합 *)
FOR _b := 1 TO GVL_PARAM.BAT_COUNT DO
	_anAuto[_b]	:= 0;
	_anManual[_b]	:= 0;
	_afBusOut[_b]	:= 0;
END_FOR
FOR _u := 1 TO GVL_PARAM.UNIT_COUNT DO
	_b := iq_astUnitCfg[_u].nBatGroup;
	IF _b >= 1 AND _b <= GVL_PARAM.BAT_COUNT THEN
		IF iq_aeOpMode[_u] = E_OpMode.Manual THEN
			_anManual[_b] := _anManual[_b] + 1;
		ELSE
			_anAuto[_b] := _anAuto[_b] + 1;
		END_IF
		IF iq_astUnit[_u].stP.bValid THEN
			_afBusOut[_b] := _afBusOut[_b] + iq_astUnit[_u].stP.fValue;
		END_IF
	END_IF
END_FOR
END_ACTION

ACTION A_CalcBusLimit:
(* 2) 버스 한도: BMS 한도 합 ∩ 버스 제한 모듈 *)
FOR _b := 1 TO GVL_PARAM.BAT_COUNT DO
	_stBatEnv	:= _stBatNone;
	_stBatEnv.stP	:= F_RangeAdd(F_RangeOpen(), F_MakeLimit(MAX(iq_astBatGroup[_b].fPDisMax, 0.0), -MAX(iq_astBatGroup[_b].fPChgMax, 0.0), GVL_REASON.RSN_BAT), 0);
	_stBatView.nBatGroup	:= _b;
	_stBatView.bUsable	:= iq_astBatGroup[_b].bUsable;
	_stBatView.stSoc	:= iq_astBatGroup[_b].stSoc;
	_stBatView.stSocMin	:= iq_astBatGroup[_b].stSocMin;
	_stBatView.stSocMax	:= iq_astBatGroup[_b].stSocMax;
	_stBatView.fPChgMax	:= iq_astBatGroup[_b].fPChgMax;
	_stBatView.fPDisMax	:= iq_astBatGroup[_b].fPDisMax;
	_stBatView.fPOut	:= _afBusOut[_b];
	_stBatView.nUnitAuto	:= _anAuto[_b];
	_stBatView.nUnitManual	:= _anManual[_b];
	FOR _i := 1 TO GVL_PARAM.BAT_RULE_COUNT DO
		IF iq_aipBatRule[_i] <> 0 AND_THEN (iq_astBatRuleReg[_i].bEnable
			AND (iq_astBatRuleReg[_i].nTarget = 0 OR iq_astBatRuleReg[_i].nTarget = _b)
			AND F_ModeApplies(iq_astBatRuleReg[_i].bAuto, iq_astBatRuleReg[_i].bManual, _anAuto[_b], _anManual[_b])) THEN
			_stBatOut	:= iq_aipBatRule[_i].M_Evaluate(_stBatView);
			_stBatEnv.stP	:= F_RangeAdd(_stBatEnv.stP, _stBatOut.stP, iq_aipBatRule[_i].ModuleId);
			_stBatEnv.bResume	:= _stBatEnv.bResume OR _stBatOut.bResume;
		END_IF
	END_FOR
	_stBatEnv.stP.fMax	:= MAX(_stBatEnv.stP.fMax, 0.0);	// 0은 항상 범위 안
	_stBatEnv.stP.fMin	:= MIN(_stBatEnv.stP.fMin, 0.0);
	q_astBatEnv[_b]	:= _stBatEnv;
END_FOR
END_ACTION

ACTION A_CalcUnitLimit:
(* 3) 유닛 한도: 정격 × Derate ∩ 유닛 제한 모듈 *)
FOR _u := 1 TO GVL_PARAM.UNIT_COUNT DO
	_stEnv	:= _stEnvNone;
	_b	:= iq_astUnitCfg[_u].nBatGroup;
	_bManual	:= iq_aeOpMode[_u] = E_OpMode.Manual;
	// 보호 상한 (P·Q 따로, 정격 대비 %). 100이면 정격
	_stEnv.bDerated	:= iq_astUnitProt[_u].fPPct < 100.0 OR iq_astUnitProt[_u].fQPct < 100.0;
	IF iq_astUnitProt[_u].fPPct < 100.0 THEN
		_fRatio	:= LIMIT(0.0, iq_astUnitProt[_u].fPPct, 100.0) / 100.0;
		_stEnv.stP	:= F_RangeAdd(F_RangeOpen(), F_MakeLimit(iq_astUnitCfg[_u].fPRated * _fRatio, -iq_astUnitCfg[_u].fPRated * _fRatio, GVL_REASON.RSN_DERATE), 0);
		_stEnv.ePMaxBy	:= E_UnitLimitBy.Derate;
		_stEnv.ePMinBy	:= E_UnitLimitBy.Derate;
	ELSE
		_stEnv.stP	:= F_RangeAdd(F_RangeOpen(), F_MakeLimit(iq_astUnitCfg[_u].fPRated, -iq_astUnitCfg[_u].fPRated, GVL_REASON.RSN_RATING), 0);
		_stEnv.ePMaxBy	:= E_UnitLimitBy.Rating;
		_stEnv.ePMinBy	:= E_UnitLimitBy.Rating;
	END_IF
	IF iq_astUnitProt[_u].fQPct < 100.0 THEN
		_fRatio	:= LIMIT(0.0, iq_astUnitProt[_u].fQPct, 100.0) / 100.0;
		_stEnv.stQ	:= F_RangeAdd(F_RangeOpen(), F_MakeLimit(iq_astUnitCfg[_u].fQRated * _fRatio, -iq_astUnitCfg[_u].fQRated * _fRatio, GVL_REASON.RSN_DERATE), 0);
		_stEnv.eQMaxBy	:= E_UnitLimitBy.Derate;
		_stEnv.eQMinBy	:= E_UnitLimitBy.Derate;
	ELSE
		_stEnv.stQ	:= F_RangeAdd(F_RangeOpen(), F_MakeLimit(iq_astUnitCfg[_u].fQRated, -iq_astUnitCfg[_u].fQRated, GVL_REASON.RSN_RATING_Q), 0);
		_stEnv.eQMaxBy	:= E_UnitLimitBy.Rating;
		_stEnv.eQMinBy	:= E_UnitLimitBy.Rating;
	END_IF
	// 피상전력 상한 = MIN(정격 S, √(P 상한² + Q 상한²)). P·Q 상한이 따로이므로 한쪽만 줄여도 다른 쪽은 묶지 않음 (둘 다 100이면 보통 정격 S)
	_fSP			:= iq_astUnitCfg[_u].fPRated * LIMIT(0.0, iq_astUnitProt[_u].fPPct, 100.0) / 100.0;
	_fSQ			:= iq_astUnitCfg[_u].fQRated * LIMIT(0.0, iq_astUnitProt[_u].fQPct, 100.0) / 100.0;
	_stEnv.fSMax	:= MIN(iq_astUnitCfg[_u].fSRated, SQRT(_fSP * _fSP + _fSQ * _fSQ));
	_stEnv.stPRule	:= F_RangeOpen();
	_stEnv.stQRule	:= F_RangeOpen();

	_stUnitView.nUnit	:= _u;
	_stUnitView.eOpMode	:= iq_aeOpMode[_u];
	_stUnitView.bAvail	:= iq_astAvail[_u].bAvail;
	_stUnitView.eRunState	:= iq_astUnit[_u].eRunState;
	_stUnitView.stP	:= iq_astUnit[_u].stP;
	_stUnitView.stQ	:= iq_astUnit[_u].stQ;
	_stUnitView.fPRated	:= iq_astUnitCfg[_u].fPRated;
	_stUnitView.fQRated	:= iq_astUnitCfg[_u].fQRated;
	_stUnitView.nBatGroup	:= _b;
	_stUnitView.stSoc	:= _stNoVal;
	IF _b >= 1 AND _b <= GVL_PARAM.BAT_COUNT THEN
		_stUnitView.stSoc := iq_astBatGroup[_b].stSoc;
	END_IF
	FOR _i := 1 TO GVL_PARAM.UNIT_RULE_COUNT DO
		IF iq_aipUnitRule[_i] <> 0 AND_THEN (iq_astUnitRuleReg[_i].bEnable
			AND (iq_astUnitRuleReg[_i].nTarget = 0 OR iq_astUnitRuleReg[_i].nTarget = _u)
			AND F_ModeApplies(iq_astUnitRuleReg[_i].bAuto, iq_astUnitRuleReg[_i].bManual, BOOL_TO_UINT(NOT _bManual), BOOL_TO_UINT(_bManual))) THEN
			_stLimOut	:= iq_aipUnitRule[_i].M_Evaluate(_stUnitView);
			_stEnv.stPRule	:= F_RangeAdd(_stEnv.stPRule, _stLimOut.stP, iq_aipUnitRule[_i].ModuleId);
			_stEnv.stQRule	:= F_RangeAdd(_stEnv.stQRule, _stLimOut.stQ, iq_aipUnitRule[_i].ModuleId);
			_stEnv.bResume	:= _stEnv.bResume OR _stLimOut.bResume;
		END_IF
	END_FOR
	// 0은 항상 범위 안 (모듈이 출력을 강제하지 못함)
	_stEnv.stPRule.fMax	:= MAX(_stEnv.stPRule.fMax, 0.0);
	_stEnv.stPRule.fMin	:= MIN(_stEnv.stPRule.fMin, 0.0);
	_stEnv.stQRule.fMax	:= MAX(_stEnv.stQRule.fMax, 0.0);
	_stEnv.stQRule.fMin	:= MIN(_stEnv.stQRule.fMin, 0.0);
	_stNew := F_RangeAnd(_stEnv.stP, _stEnv.stPRule);
	IF _stNew.fMax < _stEnv.stP.fMax THEN _stEnv.ePMaxBy := E_UnitLimitBy.UnitRule; END_IF
	IF _stNew.fMin > _stEnv.stP.fMin THEN _stEnv.ePMinBy := E_UnitLimitBy.UnitRule; END_IF
	_stEnv.stP := _stNew;
	_stNew := F_RangeAnd(_stEnv.stQ, _stEnv.stQRule);
	IF _stNew.fMax < _stEnv.stQ.fMax THEN _stEnv.eQMaxBy := E_UnitLimitBy.UnitRule; END_IF
	IF _stNew.fMin > _stEnv.stQ.fMin THEN _stEnv.eQMinBy := E_UnitLimitBy.UnitRule; END_IF
	_stEnv.stQ := _stNew;
	q_astUnitEnv[_u] := _stEnv;
END_FOR
END_ACTION

ACTION A_CalcGroupRange:
(* 4) 그룹 설비 범위 (가용 유닛). 정격 = 유닛 한도 합. 배터리 = 버스마다 min(버스 한도, 그 버스 가용 유닛 한도 합) + 배터리 없는 유닛 한도
   버스 하나를 여러 그룹이 같이 쓰면 그룹마다 버스 전체 한도를 봄 (실제 나눔은 분배가 버스 남은 한도로 맞춤) *)
FOR _g := 1 TO GVL_PARAM.GROUP_COUNT DO
	_stGrp := _stGrpNone;
	_stGrp.stRating.nMaxReason	:= GVL_REASON.RSN_RATING;
	_stGrp.stRating.nMinReason	:= GVL_REASON.RSN_RATING;
	_stGrp.stBattery.nMaxReason	:= GVL_REASON.RSN_BAT;
	_stGrp.stBattery.nMinReason	:= GVL_REASON.RSN_BAT;
	_stGrp.stQ.nMaxReason	:= GVL_REASON.RSN_RATING_Q;
	_stGrp.stQ.nMinReason	:= GVL_REASON.RSN_RATING_Q;
	FOR _b := 1 TO GVL_PARAM.BAT_COUNT DO
		_afBusMax[_b]	:= 0;
		_afBusMin[_b]	:= 0;
		_abBusIn[_b]	:= FALSE;
	END_FOR
	FOR _u := 1 TO GVL_PARAM.UNIT_COUNT DO
		IF iq_astUnitCfg[_u].nGroup = _g AND iq_astAvail[_u].bAvail THEN
			_stEnv := q_astUnitEnv[_u];
			_stGrp.stRating.fMax	:= _stGrp.stRating.fMax + _stEnv.stP.fMax;
			_stGrp.stRating.fMin	:= _stGrp.stRating.fMin + _stEnv.stP.fMin;
			_stGrp.stQ.fMax	:= _stGrp.stQ.fMax + _stEnv.stQ.fMax;
			_stGrp.stQ.fMin	:= _stGrp.stQ.fMin + _stEnv.stQ.fMin;
			_stGrp.fSMax	:= _stGrp.fSMax + _stEnv.fSMax;
			_stGrp.bResume	:= _stGrp.bResume OR _stEnv.bResume;
			// 정한 주체: 유닛 제한 모듈이 처음 찾은 것, 아니면 Derate, 아니면 정격
			IF _stGrp.stRating.nMaxModule = 0 THEN
				IF _stEnv.ePMaxBy = E_UnitLimitBy.UnitRule THEN
					_stGrp.stRating.nMaxModule	:= _stEnv.stP.nMaxModule;
					_stGrp.stRating.nMaxReason	:= _stEnv.stP.nMaxReason;
				ELSIF _stEnv.ePMaxBy = E_UnitLimitBy.Derate THEN
					_stGrp.stRating.nMaxReason	:= GVL_REASON.RSN_DERATE;
				END_IF
			END_IF
			IF _stGrp.stRating.nMinModule = 0 THEN
				IF _stEnv.ePMinBy = E_UnitLimitBy.UnitRule THEN
					_stGrp.stRating.nMinModule	:= _stEnv.stP.nMinModule;
					_stGrp.stRating.nMinReason	:= _stEnv.stP.nMinReason;
				ELSIF _stEnv.ePMinBy = E_UnitLimitBy.Derate THEN
					_stGrp.stRating.nMinReason	:= GVL_REASON.RSN_DERATE;
				END_IF
			END_IF
			_b := iq_astUnitCfg[_u].nBatGroup;
			IF _b >= 1 AND _b <= GVL_PARAM.BAT_COUNT THEN
				_afBusMax[_b]	:= _afBusMax[_b] + _stEnv.stP.fMax;
				_afBusMin[_b]	:= _afBusMin[_b] + _stEnv.stP.fMin;
				_abBusIn[_b]	:= TRUE;
			ELSE
				// 배터리 없는 유닛: 배터리 한도로 자르지 않고 자기 한도
				_stGrp.stBattery.fMax	:= _stGrp.stBattery.fMax + _stEnv.stP.fMax;
				_stGrp.stBattery.fMin	:= _stGrp.stBattery.fMin + _stEnv.stP.fMin;
			END_IF
		END_IF
	END_FOR
	FOR _b := 1 TO GVL_PARAM.BAT_COUNT DO
		IF _abBusIn[_b] THEN
			IF q_astBatEnv[_b].stP.fMax < _afBusMax[_b] THEN
				_stGrp.stBattery.fMax := _stGrp.stBattery.fMax + q_astBatEnv[_b].stP.fMax;
				IF q_astBatEnv[_b].stP.nMaxModule <> 0 AND _stGrp.stBattery.nMaxModule = 0 THEN
					_stGrp.stBattery.nMaxModule	:= q_astBatEnv[_b].stP.nMaxModule;
					_stGrp.stBattery.nMaxReason	:= q_astBatEnv[_b].stP.nMaxReason;
				END_IF
			ELSE
				_stGrp.stBattery.fMax := _stGrp.stBattery.fMax + _afBusMax[_b];
			END_IF
			IF q_astBatEnv[_b].stP.fMin > _afBusMin[_b] THEN
				_stGrp.stBattery.fMin := _stGrp.stBattery.fMin + q_astBatEnv[_b].stP.fMin;
				IF q_astBatEnv[_b].stP.nMinModule <> 0 AND _stGrp.stBattery.nMinModule = 0 THEN
					_stGrp.stBattery.nMinModule	:= q_astBatEnv[_b].stP.nMinModule;
					_stGrp.stBattery.nMinReason	:= q_astBatEnv[_b].stP.nMinReason;
				END_IF
			ELSE
				_stGrp.stBattery.fMin := _stGrp.stBattery.fMin + _afBusMin[_b];
			END_IF
			_stGrp.bResume := _stGrp.bResume OR q_astBatEnv[_b].bResume;
		END_IF
	END_FOR
	q_astGroupEnv[_g] := _stGrp;
END_FOR
END_ACTION

END_FUNCTION_BLOCK

// ---- 10_Core/40_Arbitration/F_RangeAdd.TcPOU
FUNCTION F_RangeAdd : ST_Range		// 범위를 제한 하나만큼 좁힘 (가장 좁은 범위가 남음)
VAR_INPUT
	i_stRange	: ST_Range;
	i_stLimit	: ST_Limit;
	i_nModule	: UINT;			// 제한을 낸 모듈 ID (0 = 코어)
END_VAR

F_RangeAdd := i_stRange;
IF NOT i_stLimit.bActive THEN
	RETURN;
END_IF
IF i_stLimit.fMax < F_RangeAdd.fMax THEN
	F_RangeAdd.fMax			:= i_stLimit.fMax;
	F_RangeAdd.nMaxModule	:= i_nModule;
	F_RangeAdd.nMaxReason	:= i_stLimit.nReason;
END_IF
IF i_stLimit.fMin > F_RangeAdd.fMin THEN
	F_RangeAdd.fMin			:= i_stLimit.fMin;
	F_RangeAdd.nMinModule	:= i_nModule;
	F_RangeAdd.nMinReason	:= i_stLimit.nReason;
END_IF

END_FUNCTION

// ---- 10_Core/40_Arbitration/F_RangeOpen.TcPOU
FUNCTION F_RangeOpen : ST_Range		// 제한 없는 범위
VAR
END_VAR

F_RangeOpen.fMax := 1.0E30;
F_RangeOpen.fMin := -1.0E30;

END_FUNCTION

// ---- 10_Core/40_Arbitration/F_MakeLimit.TcPOU
FUNCTION F_MakeLimit : ST_Limit		// 코어용 제한 한 줄 만들기
VAR_INPUT
	i_fMax		: REAL;
	i_fMin		: REAL;
	i_nReason	: UINT;
END_VAR

F_MakeLimit.bActive	:= TRUE;
F_MakeLimit.fMax	:= i_fMax;
F_MakeLimit.fMin	:= i_fMin;
F_MakeLimit.nReason	:= i_nReason;

END_FUNCTION

// ---- 10_Core/02_Util/F_ModeApplies.TcPOU
FUNCTION F_ModeApplies : BOOL		// 등록(bAuto·bManual)이 대상에 걸리는가: 대상 유닛 중 그 운전 모드 유닛이 하나라도 있으면. 유닛이 없는 대상(빈 버스)은 둘 중 하나라도 켜져 있으면
// 보호 조치(유닛마다)·유닛 제한·버스 제한이 같이 씀. 유닛 하나면 nAuto·nManual 중 하나만 1
VAR_INPUT
	i_bAuto		: BOOL;		// 등록: Auto 유닛에 적용
	i_bManual	: BOOL;		// 등록: Manual 유닛에 적용
	i_nAuto		: UINT;		// 대상의 Auto 유닛 수
	i_nManual	: UINT;		// 대상의 Manual 유닛 수
END_VAR

F_ModeApplies := (i_bAuto AND i_nAuto > 0) OR (i_bManual AND i_nManual > 0)
	OR (i_nAuto + i_nManual = 0 AND (i_bAuto OR i_bManual));

END_FUNCTION

// ---- 10_Core/40_Arbitration/F_RangeAnd.TcPOU
FUNCTION F_RangeAnd : ST_Range	// 두 범위의 겹치는 부분 (좁은 쪽이 이김. 상·하한마다 정한 주체를 같이 가져감)
VAR_INPUT
	i_stA	: ST_Range;
	i_stB	: ST_Range;
END_VAR

F_RangeAnd := i_stA;
IF i_stB.fMax < F_RangeAnd.fMax THEN
	F_RangeAnd.fMax	:= i_stB.fMax;
	F_RangeAnd.nMaxModule	:= i_stB.nMaxModule;
	F_RangeAnd.nMaxReason	:= i_stB.nMaxReason;
END_IF
IF i_stB.fMin > F_RangeAnd.fMin THEN
	F_RangeAnd.fMin	:= i_stB.fMin;
	F_RangeAnd.nMinModule	:= i_stB.nMinModule;
	F_RangeAnd.nMinReason	:= i_stB.nMinReason;
END_IF

END_FUNCTION

// ---- 10_Core/30_Request/FB_GroupView.TcPOU
FUNCTION_BLOCK FB_GroupView	// 제어 그룹마다 모듈에 넘길 요약을 모음 (읽기 전용)
// 가용 한도(정격·배터리)는 FB_EquipmentLimits 결과를 그대로 옮김 (여기서 다시 세지 않음). 여기서 세는 것: 정격 합(전체), 출력 합, 가용 유닛 수, SOC
VAR_IN_OUT CONSTANT
	iq_astPcc		: ARRAY[1..GVL_PARAM.GROUP_COUNT] OF ST_PccMeas;
	iq_astUnit		: ARRAY[1..GVL_PARAM.UNIT_COUNT] OF ST_UnitState;
	iq_astAvail		: ARRAY[1..GVL_PARAM.UNIT_COUNT] OF ST_UnitAvail;
	iq_astUnitCfg	: ARRAY[1..GVL_PARAM.UNIT_COUNT] OF ST_UnitCfg;
	iq_astBatGroup	: ARRAY[1..GVL_PARAM.BAT_COUNT] OF ST_BatGroupState;
	iq_aeGroupState	: ARRAY[1..GVL_PARAM.GROUP_COUNT] OF E_GroupState;	// 시퀀서 그룹 상태 (지난 스캔)
	iq_astGroupEnv	: ARRAY[1..GVL_PARAM.GROUP_COUNT] OF ST_GroupEnvelope;	// 그룹 설비 범위 (FB_EquipmentLimits)
END_VAR
VAR_OUTPUT
	q_astView		: ARRAY[1..GVL_PARAM.GROUP_COUNT] OF ST_GroupView;
END_VAR
VAR_TEMP
	g				: UINT;
	u				: UINT;
	b				: UINT;
	bSocFirst		: BOOL;
	fSocW			: REAL;
	fWSum			: REAL;
	abBatIn			: ARRAY[1..GVL_PARAM.BAT_COUNT] OF BOOL;	// 이 제어 그룹의 가용 유닛이 쓰는 배터리 그룹
	stView				: ST_GroupView;
	stNone			: ST_GroupView;
END_VAR

FOR g := 1 TO GVL_PARAM.GROUP_COUNT DO
	stView			:= stNone;
	stView.nGroup	:= g;
	stView.eState	:= iq_aeGroupState[g];
	stView.stPcc	:= iq_astPcc[g];
	FOR b := 1 TO GVL_PARAM.BAT_COUNT DO
		abBatIn[b] := FALSE;
	END_FOR

	// 유닛: 정격 합·출력 합(실측)은 전부, 가용 유닛 수
	FOR u := 1 TO GVL_PARAM.UNIT_COUNT DO
		IF iq_astUnitCfg[u].nGroup = g THEN
			stView.fPRatedSum	:= stView.fPRatedSum + iq_astUnitCfg[u].fPRated;
			stView.fQRatedSum	:= stView.fQRatedSum + iq_astUnitCfg[u].fQRated;
			IF iq_astUnit[u].stP.bValid THEN stView.fPOut := stView.fPOut + iq_astUnit[u].stP.fValue; END_IF
			IF iq_astUnit[u].stQ.bValid THEN stView.fQOut := stView.fQOut + iq_astUnit[u].stQ.fValue; END_IF
			IF iq_astAvail[u].bAvail THEN
				stView.nUnitAvail	:= stView.nUnitAvail + 1;
				b := iq_astUnitCfg[u].nBatGroup;
				IF b >= 1 AND b <= GVL_PARAM.BAT_COUNT THEN
					abBatIn[b] := TRUE;
				END_IF
			END_IF
		END_IF
	END_FOR

	// SOC: 가용 유닛이 쓰는 배터리 그룹만, 여러 유닛이 같은 그룹을 써도 한 번만 셈 (용량 가중)
	bSocFirst	:= TRUE;
	fSocW		:= 0;
	fWSum		:= 0;
	FOR b := 1 TO GVL_PARAM.BAT_COUNT DO
		IF abBatIn[b] AND iq_astBatGroup[b].bUsable THEN
			stView.fCapacity := stView.fCapacity + iq_astBatGroup[b].fCapacity;
			IF iq_astBatGroup[b].stSoc.bValid THEN
				IF bSocFirst OR iq_astBatGroup[b].stSocMin.fValue < stView.stSocMin.fValue THEN stView.stSocMin.fValue := iq_astBatGroup[b].stSocMin.fValue; END_IF
				IF bSocFirst OR iq_astBatGroup[b].stSocMax.fValue > stView.stSocMax.fValue THEN stView.stSocMax.fValue := iq_astBatGroup[b].stSocMax.fValue; END_IF
				fSocW		:= fSocW + iq_astBatGroup[b].stSoc.fValue * iq_astBatGroup[b].fSocWeight;
				fWSum		:= fWSum + iq_astBatGroup[b].fSocWeight;
				bSocFirst	:= FALSE;
			END_IF
		END_IF
	END_FOR
	IF fWSum > 0 THEN
		stView.stSocAvg.fValue	:= fSocW / fWSum;
		stView.stSocAvg.bValid	:= TRUE;
		stView.stSocMin.bValid	:= TRUE;
		stView.stSocMax.bValid	:= TRUE;
	END_IF

	// 가용 한도는 설비 한도 결과 (FB_EquipmentLimits)
	stView.fPRatedAvail	:= iq_astGroupEnv[g].stRating.fMax;
	stView.fQRatedAvail	:= iq_astGroupEnv[g].stQ.fMax;
	stView.fSRatedAvail	:= iq_astGroupEnv[g].fSMax;
	stView.fPDisMax	:= iq_astGroupEnv[g].stBattery.fMax;
	stView.fPChgMax	:= -iq_astGroupEnv[g].stBattery.fMin;
	q_astView[g] := stView;
END_FOR

END_FUNCTION_BLOCK

// ---- 10_Core/30_Request/FB_UnitView.TcPOU
FUNCTION_BLOCK FB_UnitView	// 유닛(PCS)마다 모듈에 넘길 요약 (읽기 전용). 유닛마다 제어 모드를 둘 때 씀 (FB_CtrlModeMgr.i_nUnit, MAIN이 주소를 넘김)
// 그룹 값은 FB_GroupView 결과를 받음. 여러 유닛이 한 배터리 그룹(버스)을 같이 쓰면 버스 충방전 한도·용량을 버스 가용 유닛 정격 비율로 나눔 (몫 합 = 버스 값)
// 가용이 아닌 유닛: 가용 유닛 수 0, 한도·용량·SOC 없음 (FB_GroupView가 가용 유닛만 세는 것과 같음)
VAR_IN_OUT CONSTANT
	iq_astView		: ARRAY[1..GVL_PARAM.GROUP_COUNT] OF ST_GroupView;		// FB_GroupView 결과 (이번 스캔)
	iq_astUnit		: ARRAY[1..GVL_PARAM.UNIT_COUNT] OF ST_UnitState;
	iq_astAvail		: ARRAY[1..GVL_PARAM.UNIT_COUNT] OF ST_UnitAvail;
	iq_astUnitCfg	: ARRAY[1..GVL_PARAM.UNIT_COUNT] OF ST_UnitCfg;
	iq_astUnitEnv	: ARRAY[1..GVL_PARAM.UNIT_COUNT] OF ST_UnitEnvelope;	// 유닛 한도 (FB_EquipmentLimits)
	iq_astBatGroup	: ARRAY[1..GVL_PARAM.BAT_COUNT] OF ST_BatGroupState;
	iq_astBatEnv	: ARRAY[1..GVL_PARAM.BAT_COUNT] OF ST_BatEnvelope;		// 버스 한도 (FB_EquipmentLimits)
END_VAR
VAR_OUTPUT
	q_astView		: ARRAY[1..GVL_PARAM.UNIT_COUNT] OF ST_UnitView;
END_VAR
VAR_TEMP
	u				: UINT;
	g				: UINT;
	b				: UINT;
	fShare			: REAL;
	afBusRated		: ARRAY[1..GVL_PARAM.BAT_COUNT] OF REAL;	// 버스마다 가용 유닛 정격 합
	stUv			: ST_UnitView;
	stNone			: ST_UnitView;
END_VAR

// 1) 버스마다 가용 유닛 정격 합 (버스 한도·용량을 나눌 무게)
FOR b := 1 TO GVL_PARAM.BAT_COUNT DO
	afBusRated[b] := 0;
END_FOR
FOR u := 1 TO GVL_PARAM.UNIT_COUNT DO
	b := iq_astUnitCfg[u].nBatGroup;
	IF iq_astAvail[u].bAvail AND b >= 1 AND b <= GVL_PARAM.BAT_COUNT THEN
		afBusRated[b] := afBusRated[b] + MAX(iq_astUnitCfg[u].fPRated, 0.0);
	END_IF
END_FOR

// 2) 유닛마다
FOR u := 1 TO GVL_PARAM.UNIT_COUNT DO
	stUv					:= stNone;
	stUv.nUnit				:= u;
	stUv.bAvail				:= iq_astAvail[u].bAvail;
	g						:= iq_astUnitCfg[u].nGroup;
	b						:= iq_astUnitCfg[u].nBatGroup;
	stUv.stView.nGroup		:= g;
	stUv.stView.fPRatedSum	:= iq_astUnitCfg[u].fPRated;
	stUv.stView.fQRatedSum	:= iq_astUnitCfg[u].fQRated;
	IF iq_astUnit[u].stP.bValid THEN stUv.stView.fPOut := iq_astUnit[u].stP.fValue; END_IF
	IF iq_astUnit[u].stQ.bValid THEN stUv.stView.fQOut := iq_astUnit[u].stQ.fValue; END_IF
	// 소속 그룹: 상태·접속점·출력 합
	IF g >= 1 AND g <= GVL_PARAM.GROUP_COUNT THEN
		stUv.stView.eState	:= iq_astView[g].eState;
		stUv.stView.stPcc	:= iq_astView[g].stPcc;
		stUv.fGroupPOut		:= iq_astView[g].fPOut;
		stUv.fGroupQOut		:= iq_astView[g].fQOut;
	END_IF
	IF stUv.bAvail THEN
		stUv.stView.nUnitAvail		:= 1;
		stUv.stView.fPRatedAvail	:= MAX(iq_astUnitEnv[u].stP.fMax, 0.0);
		stUv.stView.fQRatedAvail	:= MAX(iq_astUnitEnv[u].stQ.fMax, 0.0);
		stUv.stView.fSRatedAvail	:= MAX(iq_astUnitEnv[u].fSMax, 0.0);
		IF g >= 1 AND g <= GVL_PARAM.GROUP_COUNT THEN
			IF iq_astView[g].fPRatedAvail > 0 THEN
				stUv.fRatingShare := LIMIT(0.0, stUv.stView.fPRatedAvail / iq_astView[g].fPRatedAvail, 1.0);
			END_IF
		END_IF
		// 연결 버스: 한도·용량은 몫, SOC는 그대로
		IF b >= 1 AND b <= GVL_PARAM.BAT_COUNT THEN
			fShare := 0;
			IF afBusRated[b] > 0 THEN
				fShare := MAX(iq_astUnitCfg[u].fPRated, 0.0) / afBusRated[b];
			END_IF
			stUv.stView.fPDisMax	:= MIN(MAX(iq_astBatEnv[b].stP.fMax, 0.0) * fShare, stUv.stView.fPRatedAvail);
			stUv.stView.fPChgMax	:= MIN(MAX(-iq_astBatEnv[b].stP.fMin, 0.0) * fShare, stUv.stView.fPRatedAvail);
			IF iq_astBatGroup[b].bUsable THEN
				stUv.stView.fCapacity	:= iq_astBatGroup[b].fCapacity * fShare;
				stUv.stView.stSocAvg	:= iq_astBatGroup[b].stSoc;
				stUv.stView.stSocMin	:= iq_astBatGroup[b].stSocMin;
				stUv.stView.stSocMax	:= iq_astBatGroup[b].stSocMax;
			END_IF
		END_IF
	END_IF
	q_astView[u] := stUv;
END_FOR

END_FUNCTION_BLOCK

// ---- 10_Core/30_Request/FB_SourceHub.TcPOU
FUNCTION_BLOCK FB_SourceHub		// 등록된 지령원을 부르고 출력을 모음 (고르는 일은 중재에서)
VAR_IN_OUT
	iq_aipSource	: ARRAY[1..GVL_PARAM.SOURCE_COUNT] OF I_CommandSource;
END_VAR
VAR_IN_OUT CONSTANT
	iq_astReg		: ARRAY[1..GVL_PARAM.SOURCE_COUNT] OF ST_SourceReg;
	iq_astView		: ARRAY[1..GVL_PARAM.GROUP_COUNT] OF ST_GroupView;
END_VAR
VAR_OUTPUT
	q_astOut		: ARRAY[1..GVL_PARAM.SOURCE_COUNT] OF ST_SourceOutput;
	q_anModule		: ARRAY[1..GVL_PARAM.SOURCE_COUNT] OF UINT;		// 칸별 모듈 ID. 0 = 빈 칸
	q_bReset		: BOOL;			// 유효한 지령원이 PCS 리셋을 요청함 (1스캔). 유지 DO 풀기에만 씀 (장비 고장 리셋은 시퀀서가 요청을 장비별로 봄)
END_VAR
VAR_TEMP
	i				: UINT;
	g				: UINT;
	stNone			: ST_SourceOutput;
END_VAR

q_bReset := FALSE;
FOR i := 1 TO GVL_PARAM.SOURCE_COUNT DO
	IF iq_aipSource[i] <> 0 THEN
		// 대상 그룹 값을 넘김 (모든 그룹 대상이거나 번호가 틀리면 그룹 1)
		g := iq_astReg[i].nGroup;
		IF g < 1 OR g > GVL_PARAM.GROUP_COUNT THEN
			g := 1;
		END_IF
		iq_aipSource[i].M_Cycle(i_stReg := iq_astReg[i], i_stView := iq_astView[g]);
		q_astOut[i]		:= iq_aipSource[i].Output;
		q_anModule[i]	:= iq_aipSource[i].ModuleId;
	ELSE
		q_astOut[i]		:= stNone;
		q_anModule[i]	:= 0;
	END_IF

	IF q_astOut[i].bValid AND q_astOut[i].stPcsReq.eCmd = E_PcsCmd.Reset THEN
		q_bReset := TRUE;
	END_IF
END_FOR

END_FUNCTION_BLOCK

// ---- 10_Core/40_Arbitration/FB_ModeSwitch.TcPOU
FUNCTION_BLOCK FB_ModeSwitch		// 운전 모드 전환: 요청 모드 → (출력 0 → 지연 → 대기(출력 0)·정지 확인) → 실제 모드. 시작한 전환은 끝까지 진행. 보호가 ToManual을 요청하면 요청 모드를 Manual로 바꿈 (보호가 풀려도 Manual 유지)
VAR_INPUT
	i_stSet			: ST_ModeSet;
	i_fDonePct		: REAL;		// 출력 0 확인: |P|·|Q| ≤ 정격의 이 % (g_stSeqSet.stPcs.fStopDonePct, 정지 램프 완료와 같은 기준)
END_VAR
VAR_IN_OUT
	iq_aeModeReq	: ARRAY[1..GVL_PARAM.UNIT_COUNT] OF E_OpMode;		// 요청 모드 (GVL_PERSIST.g_aeOpMode). HMI가 쓰고, 보호가 ToManual을 요청하면 이 FB가 Manual로 바꿈
END_VAR
VAR_IN_OUT CONSTANT
	iq_astUnit		: ARRAY[1..GVL_PARAM.UNIT_COUNT] OF ST_UnitState;
	iq_astUnitCfg	: ARRAY[1..GVL_PARAM.UNIT_COUNT] OF ST_UnitCfg;		// 정격 (출력 0 확인)
	iq_astUnitProt	: ARRAY[1..GVL_PARAM.UNIT_COUNT] OF ST_UnitProt;	// 보호 결과 (bModeManualReq만 봄, 지난 스캔 값)
END_VAR
VAR_OUTPUT
	q_aeOpMode		: ARRAY[1..GVL_PARAM.UNIT_COUNT] OF E_OpMode;		// 실제 모드. 코어는 전부 이것을 씀
	q_abSwitching	: ARRAY[1..GVL_PARAM.UNIT_COUNT] OF BOOL;			// 전환 중: 출력 0, 지령원 상태 요청 안 받음
	q_aeStep		: ARRAY[1..GVL_PARAM.UNIT_COUNT] OF E_ModeStep;		// 진단
	q_abModeForced	: ARRAY[1..GVL_PARAM.UNIT_COUNT] OF BOOL;			// 보호가 요청 모드를 Auto에서 Manual로 바꾼 스캔 (1스캔, 기록용)
END_VAR
VAR
	_atonDelay		: ARRAY[1..GVL_PARAM.UNIT_COUNT] OF TON;
	_aeTarget		: ARRAY[1..GVL_PARAM.UNIT_COUNT] OF E_OpMode;		// 진행 중인 전환의 목표 모드 (끝날 때까지 고정)
	_bInit			: BOOL;
END_VAR
VAR_TEMP
	u				: UINT;
END_VAR

// PMS 시작: 기본은 모든 유닛 Manual로 시작 (요청 모드도 Manual로 씀). bKeepOnRestart면 저장된 요청 모드를 그대로 씀. 전환 단계 없음
// 장비 상태는 건드리지 않음: 시작 때 Run·배터리 투입 명령을 스스로 보내지 않음
IF NOT _bInit THEN
	IF NOT i_stSet.bKeepOnRestart THEN
		FOR u := 1 TO GVL_PARAM.UNIT_COUNT DO
			iq_aeModeReq[u] := E_OpMode.Manual;
		END_FOR
	END_IF
	q_aeOpMode	:= iq_aeModeReq;
	_bInit		:= TRUE;
END_IF

FOR u := 1 TO GVL_PARAM.UNIT_COUNT DO
	// 보호가 걸려 있는 동안 요청 모드는 Manual (Auto 재요청도 되돌림). 풀려도 요청은 그대로 Manual
	q_abModeForced[u] := FALSE;
	IF iq_astUnitProt[u].bModeManualReq THEN
		IF iq_aeModeReq[u] <> E_OpMode.Manual THEN
			iq_aeModeReq[u]		:= E_OpMode.Manual;
			q_abModeForced[u]	:= TRUE;
		END_IF
		// Auto로 가던 전환은 목표를 Manual로 바꿈: 끝까지 진행하는 규칙의 예외 (Auto로 한 스캔도 넘어가지 않게). 출력 0은 그대로, 남은 단계는 Manual 기준
		IF q_aeStep[u] <> E_ModeStep.Idle AND _aeTarget[u] <> E_OpMode.Manual THEN
			_aeTarget[u] := E_OpMode.Manual;
		END_IF
	END_IF
	_atonDelay[u](IN := q_aeStep[u] = E_ModeStep.Zero, PT := i_stSet.tDelay);

	IF q_aeStep[u] = E_ModeStep.Idle THEN
		// 새 전환 시작: 목표를 고정
		IF iq_aeModeReq[u] <> q_aeOpMode[u] THEN
			_aeTarget[u] := iq_aeModeReq[u];
			IF M_Level(_aeTarget[u]) = E_ModeSwitch.Direct THEN
				q_aeOpMode[u] := _aeTarget[u];
			ELSE
				q_aeStep[u] := E_ModeStep.Zero;			// 이번 스캔부터 출력 0
			END_IF
		END_IF
	ELSE
		// 진행 중: 요청이 바뀌어도 끝까지 진행. 끝난 뒤 요청이 다르면 다시 전환 (예외: 보호 ToManual은 위에서 목표를 Manual로 바꿈)
		CASE q_aeStep[u] OF
			E_ModeStep.Zero:
				IF _atonDelay[u].Q THEN
					IF M_Level(_aeTarget[u]) = E_ModeSwitch.Standby AND iq_astUnit[u].eRunState = E_RunState.Run
						AND NOT F_IsLocal(iq_astUnit[u]) THEN
						q_aeStep[u]			:= E_ModeStep.WaitStop;
					ELSE
						q_aeOpMode[u]	:= _aeTarget[u];
						q_aeStep[u]		:= E_ModeStep.Idle;
					END_IF
				END_IF

			E_ModeStep.WaitStop:
				// 대기 = 출력 0: 장비가 대기·정지를 보고하거나 실측 |P|·|Q|가 0 근처면 끝 (대기 명령은 따로 없음)
				// 로컬로 바뀌면 PMS가 제어할 수 없으므로 기다리지 않고 끝냄
				IF iq_astUnit[u].eRunState <> E_RunState.Run OR F_IsLocal(iq_astUnit[u])
					OR (ABS(iq_astUnit[u].stP.fValue) <= iq_astUnitCfg[u].fPRated * i_fDonePct / 100.0
						AND ABS(iq_astUnit[u].stQ.fValue) <= iq_astUnitCfg[u].fQRated * i_fDonePct / 100.0) THEN
					q_aeOpMode[u]	:= _aeTarget[u];
					q_aeStep[u]		:= E_ModeStep.Idle;
				END_IF
		END_CASE
	END_IF

	q_abSwitching[u] := q_aeStep[u] <> E_ModeStep.Idle;
END_FOR

METHOD PRIVATE M_Level : E_ModeSwitch		// 목표 모드로 갈 때 어디까지 하나 (MODE_SET)
VAR_INPUT
	i_eTarget	: E_OpMode;
END_VAR
IF i_eTarget = E_OpMode.Manual THEN
	M_Level := i_stSet.eToManual;
ELSE
	M_Level := i_stSet.eToAuto;
END_IF
END_METHOD

END_FUNCTION_BLOCK

// ---- 10_Core/40_Arbitration/FB_StateArbiter.TcPOU
FUNCTION_BLOCK FB_StateArbiter		// 유닛마다 이번 스캔 지령원 상태 요청 하나 고르기: 같은 스캔은 정지 쪽. 저장하지 않음 (받은 명령은 시퀀서가 한 번 보냄)
// 호출 순서 (MAIN): 본체(요청 후보) → FB_Sequencer.M_CheckRequest(접수 검사) → M_CommitRequest(접수된 것만 이번 스캔 요청)
// 보호 조치가 걸린 유닛은 그보다 기동 쪽인 요청을 버림 (보호가 풀려도 저절로 기동하지 않게). 보호 정지·비상정지 명령은 시퀀서가 보호 결과를 직접 봄
VAR_IN_OUT CONSTANT
	iq_astSrcOut	: ARRAY[1..GVL_PARAM.SOURCE_COUNT] OF ST_SourceOutput;
	iq_anSrcModule	: ARRAY[1..GVL_PARAM.SOURCE_COUNT] OF UINT;
	iq_astReg		: ARRAY[1..GVL_PARAM.SOURCE_COUNT] OF ST_SourceReg;
	iq_aeOpMode		: ARRAY[1..GVL_PARAM.UNIT_COUNT] OF E_OpMode;
	iq_astUnitCfg	: ARRAY[1..GVL_PARAM.UNIT_COUNT] OF ST_UnitCfg;
	iq_astUnitProt	: ARRAY[1..GVL_PARAM.UNIT_COUNT] OF ST_UnitProt;
	iq_abSwitching	: ARRAY[1..GVL_PARAM.UNIT_COUNT] OF BOOL;		// 모드 전환 중: 지령원 기동 쪽 요청(Run) 안 받음. 정지 쪽은 받음
END_VAR
VAR_OUTPUT
	(* 요청 후보 (본체 결과, 접수 검사 전) *)
	q_abCand		: ARRAY[1..GVL_PARAM.UNIT_COUNT] OF BOOL;		// 이번 스캔 요청 후보 있음
	q_aeCand		: ARRAY[1..GVL_PARAM.UNIT_COUNT] OF E_PcsCmd;	// 후보 명령
	q_anCandModule	: ARRAY[1..GVL_PARAM.UNIT_COUNT] OF UINT;		// 후보를 낸 지령원 모듈 ID
	(* 이번 스캔 요청 (M_CommitRequest 결과) *)
	q_abNewReq		: ARRAY[1..GVL_PARAM.UNIT_COUNT] OF BOOL;		// 이번 스캔에 접수된 요청 있음
	q_aeReq			: ARRAY[1..GVL_PARAM.UNIT_COUNT] OF E_PcsCmd;	// 그 요청 (없으면 None)
	q_abPcsReqTaken	: ARRAY[1..GVL_PARAM.SOURCE_COUNT] OF BOOL;		// 지령원의 이번 PCS 요청을 후보로 본 유닛이 있음 (로그용. FALSE면 운전 모드 설정·모드 전환 때문에 무시)
END_VAR
VAR_TEMP
	u				: UINT;
	i				: UINT;
	nRank			: INT;
	nBest			: INT;
	eBest			: E_PcsCmd;
	nBestModule		: UINT;
	nProtRank		: INT;
END_VAR

FOR i := 1 TO GVL_PARAM.SOURCE_COUNT DO
	q_abPcsReqTaken[i] := FALSE;
END_FOR
FOR u := 1 TO GVL_PARAM.UNIT_COUNT DO
	// 1) 이번 스캔 요청 중 가장 정지 쪽 (이 유닛의 운전 모드에 맞는 지령원만)
	nBest		:= -1;
	eBest		:= E_PcsCmd.None;
	nBestModule	:= 0;
	FOR i := 1 TO GVL_PARAM.SOURCE_COUNT DO
		nRank := F_StateRank(iq_astSrcOut[i].stPcsReq.eCmd);
		IF iq_astSrcOut[i].bValid AND nRank >= 0
			AND (iq_astReg[i].nGroup = 0 OR iq_astReg[i].nGroup = iq_astUnitCfg[u].nGroup)
			AND (iq_astSrcOut[i].stPcsReq.nUnit = 0 OR iq_astSrcOut[i].stPcsReq.nUnit = u)
			AND F_PcsCmdAllowed(iq_astReg[i].stStateMode.stPcs, iq_astSrcOut[i].stPcsReq.eCmd, iq_aeOpMode[u])
			AND (NOT iq_abSwitching[u] OR nRank >= F_StateRank(E_PcsCmd.Standby)) THEN		// 모드 전환 중에는 정지 쪽(Standby·Stop·EStop)만 받음
			q_abPcsReqTaken[i] := TRUE;
			IF nRank > nBest THEN
				nBest		:= nRank;
				eBest		:= iq_astSrcOut[i].stPcsReq.eCmd;
				nBestModule	:= iq_anSrcModule[i];
			END_IF
		END_IF
	END_FOR
	// 2) 보호 조치보다 기동 쪽인 요청은 버림 (접수 검사 전)
	CASE iq_astUnitProt[u].ePcsAction OF
		E_PcsAction.Standby:	nProtRank := F_StateRank(E_PcsCmd.Standby);
		E_PcsAction.Stop:		nProtRank := F_StateRank(E_PcsCmd.Stop);
		E_PcsAction.EStop:		nProtRank := F_StateRank(E_PcsCmd.EStop);
	ELSE
		nProtRank := -1;
	END_CASE
	q_abCand[u]			:= nBest >= 0 AND nBest >= nProtRank;
	q_aeCand[u]			:= eBest;
	q_anCandModule[u]	:= nBestModule;
	q_abNewReq[u]		:= FALSE;		// M_CommitRequest에서 정함
	q_aeReq[u]			:= E_PcsCmd.None;
END_FOR

METHOD M_CommitRequest		// 접수된 후보만 이번 스캔 요청으로 (거부된 후보는 버림)
VAR_IN_OUT CONSTANT
	iq_abAccept		: ARRAY[1..GVL_PARAM.UNIT_COUNT] OF BOOL;		// 접수 검사 결과 (FB_Sequencer.q_abAccept)
END_VAR
VAR
	u				: UINT;
END_VAR
FOR u := 1 TO GVL_PARAM.UNIT_COUNT DO
	q_abNewReq[u] := q_abCand[u] AND iq_abAccept[u];
	IF q_abNewReq[u] THEN
		q_aeReq[u] := q_aeCand[u];
	END_IF
END_FOR
END_METHOD

END_FUNCTION_BLOCK

// ---- 10_Core/40_Arbitration/F_StateRank.TcPOU
FUNCTION F_StateRank : INT		// 상태 요청 세기 (정지 쪽이 큼). 상태가 아닌 요청은 -1
VAR_INPUT
	i_eCmd		: E_PcsCmd;
END_VAR

CASE i_eCmd OF
	E_PcsCmd.Run:		F_StateRank := 0;
	E_PcsCmd.Standby:	F_StateRank := 1;
	E_PcsCmd.Stop:	F_StateRank := 2;
	E_PcsCmd.EStop:	F_StateRank := 3;
ELSE
	F_StateRank := -1;		// None, Reset
END_CASE

END_FUNCTION

// ---- 10_Core/40_Arbitration/F_PcsCmdAllowed.TcPOU
FUNCTION F_PcsCmdAllowed : BOOL		// 지령원의 PCS 요청을 이 운전 모드에서 받나 (명령마다 등록값). 리셋은 항상 받음
VAR_INPUT
	i_stSet		: ST_PcsCmdMode;
	i_eCmd		: E_PcsCmd;
	i_eOpMode	: E_OpMode;
END_VAR

CASE i_eCmd OF
	E_PcsCmd.Run:		F_PcsCmdAllowed := F_SourceAllowed(i_stSet.eRun, i_eOpMode);
	E_PcsCmd.Standby:	F_PcsCmdAllowed := F_SourceAllowed(i_stSet.eStandby, i_eOpMode);
	E_PcsCmd.Stop:		F_PcsCmdAllowed := F_SourceAllowed(i_stSet.eStop, i_eOpMode);
	E_PcsCmd.EStop:		F_PcsCmdAllowed := F_SourceAllowed(i_stSet.eEStop, i_eOpMode);
	E_PcsCmd.Reset:		F_PcsCmdAllowed := TRUE;
ELSE
	F_PcsCmdAllowed := FALSE;		// None
END_CASE

END_FUNCTION

// ---- 10_Core/40_Arbitration/F_SourceAllowed.TcPOU
FUNCTION F_SourceAllowed : BOOL		// 지령원이 이 운전 모드에서 동작하나
VAR_INPUT
	i_eSrcMode	: E_SourceMode;
	i_eOpMode	: E_OpMode;
END_VAR

CASE i_eSrcMode OF
	E_SourceMode.Both:		F_SourceAllowed := TRUE;
	E_SourceMode.Auto:		F_SourceAllowed := (i_eOpMode = E_OpMode.Auto);
	E_SourceMode.Manual:	F_SourceAllowed := (i_eOpMode = E_OpMode.Manual);
ELSE
	F_SourceAllowed := FALSE;
END_CASE

END_FUNCTION

// ---- 10_Core/40_Arbitration/FB_Select.TcPOU
FUNCTION_BLOCK FB_Select		// 지령원 중에서 유닛별 값과 그룹 값을 고름 (지령원 P·Q 제한은 모두 겹침). Auto 경로·Manual 경로로 나눠 냄 (고르는 규칙은 같음)
// 이상값을 뺀 후보를 고르기 정책(그룹마다 I_SelectPolicy, 비우면 코어 기본 FB_SelectStd)에 넘김. 정책이 낸 값도 이상값이면 버림
VAR_IN_OUT
	iq_aipSelPolicy	: ARRAY[1..GVL_PARAM.GROUP_COUNT] OF I_SelectPolicy;	// 그룹별 고르기 정책 (GVL_SITE.g_aipSelectPolicy)
END_VAR
VAR_IN_OUT CONSTANT
	iq_astSrcOut	: ARRAY[1..GVL_PARAM.SOURCE_COUNT] OF ST_SourceOutput;
	iq_anSrcModule	: ARRAY[1..GVL_PARAM.SOURCE_COUNT] OF UINT;
	iq_astReg		: ARRAY[1..GVL_PARAM.SOURCE_COUNT] OF ST_SourceReg;
	iq_aeOpMode		: ARRAY[1..GVL_PARAM.UNIT_COUNT] OF E_OpMode;
	iq_astUnitCfg	: ARRAY[1..GVL_PARAM.UNIT_COUNT] OF ST_UnitCfg;
	iq_astGroupSet	: ARRAY[1..GVL_PARAM.GROUP_COUNT] OF ST_GroupSet;
	iq_astView		: ARRAY[1..GVL_PARAM.GROUP_COUNT] OF ST_GroupView;	// 그룹 유닛 정격 합 (이상값 한도)
	iq_stFilter		: ST_CmdFilterSet;
END_VAR
VAR_OUTPUT
	(* Auto 경로 *)
	q_astAutoUnitP	: ARRAY[1..GVL_PARAM.UNIT_COUNT] OF ST_Pick;		// Auto 유닛의 유닛별 P 값 (kW, 유닛 출력). Manual 유닛은 비활성
	q_astAutoUnitQ	: ARRAY[1..GVL_PARAM.UNIT_COUNT] OF ST_Pick;
	q_astAutoGrpP	: ARRAY[1..GVL_PARAM.GROUP_COUNT] OF ST_Pick;		// kW, 접속점 기준
	q_astAutoGrpQ	: ARRAY[1..GVL_PARAM.GROUP_COUNT] OF ST_Pick;
	q_astAutoGrpPLim: ARRAY[1..GVL_PARAM.GROUP_COUNT] OF ST_Range;		// Auto 지령원들이 낸 P 제한 (접속점 기준)
	(* Manual 경로 *)
	q_astManualUnitP: ARRAY[1..GVL_PARAM.UNIT_COUNT] OF ST_Pick;		// Manual 유닛의 유닛별 P 값. Auto 유닛은 비활성
	q_astManualUnitQ: ARRAY[1..GVL_PARAM.UNIT_COUNT] OF ST_Pick;
	q_astManualGrpP	: ARRAY[1..GVL_PARAM.GROUP_COUNT] OF ST_Pick;		// kW, 그룹 값 (그룹의 Manual 유닛에 나눔)
	q_astManualGrpQ	: ARRAY[1..GVL_PARAM.GROUP_COUNT] OF ST_Pick;
	q_astManualGrpPLim: ARRAY[1..GVL_PARAM.GROUP_COUNT] OF ST_Range;	// Manual 지령원들이 낸 P 제한
	q_astAutoGrpQLim: ARRAY[1..GVL_PARAM.GROUP_COUNT] OF ST_Range;		// Auto 지령원들이 낸 Q 제한 (접속점 기준)
	q_astManualGrpQLim: ARRAY[1..GVL_PARAM.GROUP_COUNT] OF ST_Range;	// Manual 지령원들이 낸 Q 제한
	(* 이상값으로 무시한 지령원 *)
	q_abBadValue	: ARRAY[1..GVL_PARAM.SOURCE_COUNT] OF BOOL;		// 이번 스캔에 이상값이 있었음
	q_afBadValue	: ARRAY[1..GVL_PARAM.SOURCE_COUNT] OF REAL;		// 그 값 (진단용)
	q_anPolicyBad	: UINT;		// 이번 스캔에 정책이 이상값을 내 버린 수 (진단)
END_VAR
VAR
	_fbSelStd		: FB_SelectStd;		// 코어 기본 고르기 정책
	_aipSelPolicy	: ARRAY[1..GVL_PARAM.GROUP_COUNT] OF I_SelectPolicy;	// 사본 (메서드에서 씀)
END_VAR
VAR_TEMP
	u				: UINT;
	g				: UINT;
	i				: UINT;
	k				: UINT;
	eMode			: E_OpMode;
	stPickP			: ST_Pick;
	stPickQ			: ST_Pick;
	stViewP			: ST_SelectView;	// 고르기 후보 (P)
	stViewQ			: ST_SelectView;
	stViewNone		: ST_SelectView;
	stRng			: ST_Range;		// 지령원 P 제한 모음
	stQRng			: ST_Range;		// 지령원 Q 제한 모음
	stLim			: ST_Limit;
	stNone			: ST_Pick;
	fLimP			: REAL;			// 이상값 한도 (0 = 검사 안 함)
	fLimQ			: REAL;
	stUnitP			: ST_Pick;		// 이번 유닛에서 고른 값 (운전 모드에 맞는 경로로 보냄)
	stUnitQ			: ST_Pick;
END_VAR

_aipSelPolicy := iq_aipSelPolicy;
q_anPolicyBad := 0;
(* 0) 이상값 한도 준비 *)
FOR i := 1 TO GVL_PARAM.SOURCE_COUNT DO
	q_abBadValue[i] := FALSE;
END_FOR

(* 1) 유닛별 값: 이 유닛의 운전 모드에 맞는 지령원 후보 (이상값은 뺌) → 정책 (기본: 등급이 가장 높은 것) *)
FOR u := 1 TO GVL_PARAM.UNIT_COUNT DO
	stViewP			:= stViewNone;
	stViewP.nGroup	:= iq_astUnitCfg[u].nGroup;
	stViewP.nUnit	:= u;
	stViewP.eOpMode	:= iq_aeOpMode[u];
	stViewQ			:= stViewP;
	stViewQ.bForQ	:= TRUE;
	fLimP			:= SEL(iq_stFilter.bBadValue, 0.0, iq_astUnitCfg[u].fPRated * iq_stFilter.fBadFactor);
	fLimQ			:= SEL(iq_stFilter.bBadValue, 0.0, iq_astUnitCfg[u].fQRated * iq_stFilter.fBadFactor);
	FOR i := 1 TO GVL_PARAM.SOURCE_COUNT DO
		IF iq_astSrcOut[i].bValid
			AND (iq_astReg[i].nGroup = 0 OR iq_astReg[i].nGroup = iq_astUnitCfg[u].nGroup)
			AND F_SourceAllowed(iq_astReg[i].ePowerMode, iq_aeOpMode[u]) THEN
			IF iq_astSrcOut[i].astUnit[u].bPSetActive AND NOT F_CmdOk(iq_astSrcOut[i].astUnit[u].fPSet, fLimP) THEN
				q_abBadValue[i] := TRUE;
				q_afBadValue[i] := iq_astSrcOut[i].astUnit[u].fPSet;
			ELSIF iq_astSrcOut[i].astUnit[u].bPSetActive THEN
				M_AddCand(stViewP, i, iq_anSrcModule[i], iq_astReg[i].nGrade, iq_astSrcOut[i].astUnit[u].fPSet, iq_astSrcOut[i].bNewSet);
			END_IF
			IF iq_astSrcOut[i].astUnit[u].bQSetActive AND NOT F_CmdOk(iq_astSrcOut[i].astUnit[u].fQSet, fLimQ) THEN
				q_abBadValue[i] := TRUE;
				q_afBadValue[i] := iq_astSrcOut[i].astUnit[u].fQSet;
			ELSIF iq_astSrcOut[i].astUnit[u].bQSetActive THEN
				M_AddCand(stViewQ, i, iq_anSrcModule[i], iq_astReg[i].nGrade, iq_astSrcOut[i].astUnit[u].fQSet, iq_astSrcOut[i].bNewSet);
			END_IF
		END_IF
	END_FOR
	stUnitP := M_Pick(stViewP, fLimP);
	stUnitQ := M_Pick(stViewQ, fLimQ);
	// 운전 모드에 맞는 경로로
	q_astAutoUnitP[u]	:= stNone;
	q_astAutoUnitQ[u]	:= stNone;
	q_astManualUnitP[u]	:= stNone;
	q_astManualUnitQ[u]	:= stNone;
	IF iq_aeOpMode[u] = E_OpMode.Manual THEN
		q_astManualUnitP[u]	:= stUnitP;
		q_astManualUnitQ[u]	:= stUnitQ;
	ELSE
		q_astAutoUnitP[u]	:= stUnitP;
		q_astAutoUnitQ[u]	:= stUnitQ;
	END_IF
END_FOR

(* 2) 그룹 값: 운전 모드(Auto / Manual)마다 따로 후보를 모아 정책으로 고름 (기본: eSelP·eSelQ). 지령원 P·Q 제한은 모두 모음 *)
FOR g := 1 TO GVL_PARAM.GROUP_COUNT DO
	FOR k := 1 TO 2 DO
		IF k = 1 THEN
			eMode := E_OpMode.Auto;
		ELSE
			eMode := E_OpMode.Manual;
		END_IF
		stViewP			:= stViewNone;
		stViewP.nGroup	:= g;
		stViewP.eOpMode	:= eMode;
		stViewP.eSel	:= iq_astGroupSet[g].eSelP;
		stViewQ			:= stViewP;
		stViewQ.bForQ	:= TRUE;
		stViewQ.eSel	:= iq_astGroupSet[g].eSelQ;
		stRng	:= F_RangeOpen();
		stQRng	:= F_RangeOpen();
		fLimP	:= SEL(iq_stFilter.bBadValue, 0.0, iq_astView[g].fPRatedSum * iq_stFilter.fBadFactor);
		fLimQ	:= SEL(iq_stFilter.bBadValue, 0.0, iq_astView[g].fQRatedSum * iq_stFilter.fBadFactor);

		FOR i := 1 TO GVL_PARAM.SOURCE_COUNT DO
			IF iq_astSrcOut[i].bValid
				AND (iq_astReg[i].nGroup = 0 OR iq_astReg[i].nGroup = g)
				AND F_SourceAllowed(iq_astReg[i].ePowerMode, eMode) THEN
				IF iq_astSrcOut[i].bPSetActive AND NOT F_CmdOk(iq_astSrcOut[i].fPSet, fLimP) THEN
					q_abBadValue[i] := TRUE;
					q_afBadValue[i] := iq_astSrcOut[i].fPSet;
				ELSIF iq_astSrcOut[i].bPSetActive THEN
					M_AddCand(stViewP, i, iq_anSrcModule[i], iq_astReg[i].nGrade, iq_astSrcOut[i].fPSet, iq_astSrcOut[i].bNewSet);
				END_IF
				IF iq_astSrcOut[i].bQSetActive AND NOT F_CmdOk(iq_astSrcOut[i].fQSet, fLimQ) THEN
					q_abBadValue[i] := TRUE;
					q_afBadValue[i] := iq_astSrcOut[i].fQSet;
				ELSIF iq_astSrcOut[i].bQSetActive THEN
					M_AddCand(stViewQ, i, iq_anSrcModule[i], iq_astReg[i].nGrade, iq_astSrcOut[i].fQSet, iq_astSrcOut[i].bNewSet);
				END_IF
				// [결함 13 수정 2026-11-04: 지령원 P·Q 제한값이 숫자가 아니면 이상값으로 보고 그 제한은 안 씀 (범위 계산 비교에서 FPU 예외)]
				IF iq_astSrcOut[i].bPLimActive AND NOT (F_RealOk(iq_astSrcOut[i].fPMax) AND F_RealOk(iq_astSrcOut[i].fPMin)) THEN
					q_abBadValue[i] := TRUE;
					q_afBadValue[i] := SEL(F_RealOk(iq_astSrcOut[i].fPMax), iq_astSrcOut[i].fPMax, iq_astSrcOut[i].fPMin);
				ELSIF iq_astSrcOut[i].bPLimActive THEN
					stLim.bActive	:= TRUE;
					stLim.fMax		:= iq_astSrcOut[i].fPMax;
					stLim.fMin		:= iq_astSrcOut[i].fPMin;
					stLim			:= F_LimitKeepZero(stLim);		// 0은 항상 범위 안
					stLim.nReason	:= 0;
					stRng := F_RangeAdd(stRng, stLim, iq_anSrcModule[i]);
				END_IF
				IF iq_astSrcOut[i].bQLimActive AND NOT (F_RealOk(iq_astSrcOut[i].fQMax) AND F_RealOk(iq_astSrcOut[i].fQMin)) THEN	// [결함 13 수정 2026-11-04]
					q_abBadValue[i] := TRUE;
					q_afBadValue[i] := SEL(F_RealOk(iq_astSrcOut[i].fQMax), iq_astSrcOut[i].fQMax, iq_astSrcOut[i].fQMin);
				ELSIF iq_astSrcOut[i].bQLimActive THEN
					stLim.bActive	:= TRUE;
					stLim.fMax		:= iq_astSrcOut[i].fQMax;
					stLim.fMin		:= iq_astSrcOut[i].fQMin;
					stLim			:= F_LimitKeepZero(stLim);
					stLim.nReason	:= 0;
					stQRng := F_RangeAdd(stQRng, stLim, iq_anSrcModule[i]);
				END_IF
			END_IF
		END_FOR

		stPickP := M_Pick(stViewP, fLimP);
		stPickQ := M_Pick(stViewQ, fLimQ);
		IF k = 1 THEN
			q_astAutoGrpP[g]		:= stPickP;
			q_astAutoGrpQ[g]		:= stPickQ;
			q_astAutoGrpPLim[g]		:= stRng;
			q_astAutoGrpQLim[g]		:= stQRng;
		ELSE
			q_astManualGrpP[g]		:= stPickP;
			q_astManualGrpQ[g]		:= stPickQ;
			q_astManualGrpPLim[g]	:= stRng;
			q_astManualGrpQLim[g]	:= stQRng;
		END_IF
	END_FOR
END_FOR

METHOD PRIVATE M_AddCand		// 후보 하나 추가 (지령원 칸 순서)
VAR_IN_OUT
	iq_stView	: ST_SelectView;
END_VAR
VAR_INPUT
	i_nSource	: UINT;
	i_nModule	: UINT;
	i_nGrade	: UINT;
	i_fValue	: REAL;
	i_bNew		: BOOL;
END_VAR
IF iq_stView.nCand >= GVL_PARAM.SOURCE_COUNT THEN
	RETURN;
END_IF
iq_stView.nCand := iq_stView.nCand + 1;
iq_stView.astCand[iq_stView.nCand].nSource	:= i_nSource;
iq_stView.astCand[iq_stView.nCand].nModule	:= i_nModule;
iq_stView.astCand[iq_stView.nCand].nGrade	:= i_nGrade;
iq_stView.astCand[iq_stView.nCand].fValue	:= i_fValue;
iq_stView.astCand[iq_stView.nCand].bNew		:= i_bNew;
END_METHOD

METHOD PRIVATE M_Pick : ST_Pick		// 후보를 정책에 넘겨 하나로. 그룹에 정책이 없으면 코어 기본. 후보가 없으면 값 없음, 정책이 낸 값이 이상값이면 버림
VAR_INPUT
	i_stView	: ST_SelectView;
	i_fLim		: REAL;			// 이상값 한도 (0 = 크기 검사 안 함)
END_VAR
IF i_stView.nCand = 0 THEN
	RETURN;
END_IF
IF i_stView.nGroup >= 1 AND i_stView.nGroup <= GVL_PARAM.GROUP_COUNT AND_THEN _aipSelPolicy[i_stView.nGroup] <> 0 THEN
	M_Pick := _aipSelPolicy[i_stView.nGroup].M_Select(i_stView := i_stView);
ELSE
	M_Pick := _fbSelStd.M_Select(i_stView := i_stView);
END_IF
IF M_Pick.bActive AND NOT F_CmdOk(M_Pick.fValue, i_fLim) THEN
	M_Pick.bActive	:= FALSE;
	q_anPolicyBad	:= q_anPolicyBad + 1;
END_IF
END_METHOD

END_FUNCTION_BLOCK

// ---- 10_Core/40_Arbitration/FB_SelectStd.TcPOU
FUNCTION_BLOCK FB_SelectStd EXTENDS FB_ModuleBase IMPLEMENTS I_SelectPolicy	// 코어 기본 고르기: 유닛별 값은 등급, 그룹 값은 그룹 설정 eSelP·eSelQ (등급 / 절대값 작은 것). 같으면 먼저 등록된 칸

METHOD M_Select : ST_Pick
VAR_INPUT
	i_stView	: ST_SelectView;
END_VAR
VAR
	i		: UINT;
	eSel	: E_SelectMode;
	nGrade	: UINT;
END_VAR
eSel := E_SelectMode.Grade;		// 유닛별 값은 등급만
IF i_stView.nUnit = 0 THEN
	eSel := i_stView.eSel;
END_IF
FOR i := 1 TO MIN(i_stView.nCand, GVL_PARAM.SOURCE_COUNT) DO
	IF F_Better(eSel, M_Select.bActive, i_stView.astCand[i].nGrade, i_stView.astCand[i].fValue, nGrade, M_Select.fValue) THEN
		M_Select.bActive	:= TRUE;
		M_Select.fValue		:= i_stView.astCand[i].fValue;
		M_Select.nModule	:= i_stView.astCand[i].nModule;
		M_Select.bNew		:= i_stView.astCand[i].bNew;
		nGrade				:= i_stView.astCand[i].nGrade;
	END_IF
END_FOR
END_METHOD

END_FUNCTION_BLOCK

// ---- 10_Core/03_Base/FB_ModuleBase.TcPOU
FUNCTION_BLOCK ABSTRACT FB_ModuleBase IMPLEMENTS I_Module
VAR_INPUT
	i_nModuleId		: UINT;			// 현장 안에서 겹치지 않는 번호. GVL_SITE에서 정함
	i_sName			: STRING(31);	// 로그에 나오는 이름 (영문)
END_VAR

PROPERTY ModuleId : UINT
GET
ModuleId := i_nModuleId;
END_GET
END_PROPERTY

PROPERTY ModuleName : STRING(31)
GET
ModuleName := i_sName;
END_GET
END_PROPERTY

METHOD M_ReasonText : WSTRING(63)		// 기본: "이유 n". 모듈이 바꿔서 자기 문구를 돌려줌
VAR_INPUT
	i_nReason	: UINT;
END_VAR
M_ReasonText := WCONCAT("이유 ", TO_WSTRING(i_nReason));
END_METHOD

METHOD M_CheckSet : WSTRING(63)		// 기본: 점검할 설정 없음 (빈 문구). 설정 구조체를 받는 모듈이 바꿔서 자기 설정을 점검
M_CheckSet := "";
END_METHOD

END_FUNCTION_BLOCK

// ---- 10_Core/40_Arbitration/F_Better.TcPOU
FUNCTION F_Better : BOOL		// 새 후보가 지금 고른 것보다 나은가
VAR_INPUT
	i_eSel		: E_SelectMode;
	i_bHave		: BOOL;			// 이미 고른 것이 있음
	i_nGrade	: UINT;			// 새 후보 등급
	i_fValue	: REAL;
	i_nGradeOld	: UINT;
	i_fValueOld	: REAL;
END_VAR

IF NOT i_bHave THEN
	F_Better := TRUE;
ELSIF i_eSel = E_SelectMode.MinAbs AND ABS(i_fValue) <> ABS(i_fValueOld) THEN
	F_Better := ABS(i_fValue) < ABS(i_fValueOld);
ELSE
	F_Better := i_nGrade < i_nGradeOld;		// 같으면 먼저 등록된 칸 유지
END_IF

END_FUNCTION

// ---- 10_Core/02_Util/F_RealOk.TcPOU
FUNCTION F_RealOk : BOOL		// REAL이 숫자인가 (NaN·±무한대면 FALSE). 비교하지 않고 비트로 봄 → FPU 예외 없음 [결함 13 수정 2026-11-04: 추가]
// TwinCAT x86/x64는 FPU 예외가 켜져 있어 NaN을 비교(=, <, <=)·변환(REAL_TO_*, LIMIT)하면 PLC가 멈춤. 밖에서 들어온 REAL은 쓰기 전에 이 함수로 먼저 거름
// (Tc2_Utilities.IsFinite(F_REAL(x))와 같은 판단. 코어 함수라 라이브러리에 기대지 않음)
VAR_INPUT
	i_fValue	: REAL;
END_VAR
VAR
	dwBits		: DWORD;
END_VAR

MEMCPY(ADR(dwBits), ADR(i_fValue), SIZEOF(dwBits));
F_RealOk := (dwBits AND 16#7F800000) <> 16#7F800000;	// 지수 8비트가 모두 1 = NaN 또는 ±무한대

END_FUNCTION

// ---- 10_Core/40_Arbitration/F_LimitKeepZero.TcPOU
FUNCTION F_LimitKeepZero : ST_Limit		// 제한은 줄이기만 함: 0은 항상 범위 안 (상한 < 0, 하한 > 0이면 0으로. 강제 출력은 지령으로). NaN은 그대로 (F_Range가 무시)
VAR_INPUT
	i_stLim		: ST_Limit;
END_VAR

F_LimitKeepZero := i_stLim;
IF F_LimitKeepZero.fMax < 0.0 THEN F_LimitKeepZero.fMax := 0.0; END_IF
IF F_LimitKeepZero.fMin > 0.0 THEN F_LimitKeepZero.fMin := 0.0; END_IF

END_FUNCTION

// ---- 10_Core/40_Arbitration/FB_Gate.TcPOU
FUNCTION_BLOCK FB_Gate		// 경로별 지령 거르기 자리 (Auto·Manual이 같은 FB를 경로만 바꿔 두 번 씀): 등록한 Gate 모듈(i_ipGate), 비우면 그 경로의 코어 기본 Gate. 출력 모양은 고정 (뒤 단계는 이것만 봄)
// 뒤 단계(성형·분배·보호·쓰기 허가)는 Gate와 관계없이 그대로 적용됨
VAR_INPUT
	i_ePath			: E_OpMode;			// 이 인스턴스가 맡는 경로 (Auto 또는 Manual)
	i_ipGate		: I_Gate;			// GVL_SITE.g_ipAutoGate·g_ipManualGate. 0 = 그 경로의 코어 기본 (Auto = FB_GateAuto, Manual = FB_GateManual)
	i_stManualCmdSet	: ST_ManualCmdSet;	// Manual 지령 거르기 설정 (코어 기본 Manual Gate가 씀. Auto 경로는 연결하지 않음)
END_VAR
VAR_IN_OUT CONSTANT
	iq_astUnitP		: ARRAY[1..GVL_PARAM.UNIT_COUNT] OF ST_Pick;		// 이 경로 FB_Select 결과
	iq_astUnitQ		: ARRAY[1..GVL_PARAM.UNIT_COUNT] OF ST_Pick;
	iq_astGrpP		: ARRAY[1..GVL_PARAM.GROUP_COUNT] OF ST_Pick;
	iq_astGrpQ		: ARRAY[1..GVL_PARAM.GROUP_COUNT] OF ST_Pick;
	iq_aeOpMode		: ARRAY[1..GVL_PARAM.UNIT_COUNT] OF E_OpMode;
	iq_astUnit		: ARRAY[1..GVL_PARAM.UNIT_COUNT] OF ST_UnitState;
	iq_astUnitCfg	: ARRAY[1..GVL_PARAM.UNIT_COUNT] OF ST_UnitCfg;
END_VAR
VAR_OUTPUT
	(* 거른 결과: 성형·분배는 이것을 씀 *)
	q_astUnitP		: ARRAY[1..GVL_PARAM.UNIT_COUNT] OF ST_Pick;
	q_astUnitQ		: ARRAY[1..GVL_PARAM.UNIT_COUNT] OF ST_Pick;
	q_astGrpP		: ARRAY[1..GVL_PARAM.GROUP_COUNT] OF ST_Pick;
	q_astGrpQ		: ARRAY[1..GVL_PARAM.GROUP_COUNT] OF ST_Pick;
	q_abNew			: ARRAY[1..GVL_PARAM.UNIT_COUNT] OF BOOL;			// 새 지령을 받아들임 (Manual 경로: 디스패처가 이 스캔에 바로 씀)
	(* 진단 *)
	q_aeRefuse		: ARRAY[1..GVL_PARAM.UNIT_COUNT] OF E_CmdRefuse;		// 마지막으로 무시한 이유 (새 지령을 받아들이면 None)
	q_anRefuseModule: ARRAY[1..GVL_PARAM.UNIT_COUNT] OF UINT;			// 무시한 지령을 낸 모듈 ID
	q_abWaitNewCmd	: ARRAY[1..GVL_PARAM.UNIT_COUNT] OF BOOL;			// Manual 유닛: Run 확인 뒤 새 지령이 올 때까지 출력 0
END_VAR
VAR
	_fbAuto		: FB_GateAuto;		// 코어 기본 Auto Gate
	_fbManual	: FB_GateManual;	// 코어 기본 Manual Gate
	_ipUse		: I_Gate;			// 이번 스캔에 쓰는 Gate
	_stOut		: ST_GateOut;
END_VAR
VAR_TEMP
	u			: UINT;
	stView		: ST_GateView;
	stNone		: ST_Pick;
	bManualPath	: BOOL;
END_VAR

bManualPath		:= i_ePath = E_OpMode.Manual;
stView.ePath		:= i_ePath;
stView.stManualCmdSet	:= i_stManualCmdSet;

// 쓸 Gate: 등록한 모듈, 없으면 이 경로의 코어 기본
_ipUse := i_ipGate;
IF _ipUse = 0 THEN
	IF bManualPath THEN
		_ipUse := _fbManual;
	ELSE
		_ipUse := _fbAuto;
	END_IF
END_IF
_ipUse.M_Filter(i_stView := stView, iq_astUnitP := iq_astUnitP, iq_astUnitQ := iq_astUnitQ, iq_astGrpP := iq_astGrpP, iq_astGrpQ := iq_astGrpQ,
	iq_aeOpMode := iq_aeOpMode, iq_astUnit := iq_astUnit, iq_astUnitCfg := iq_astUnitCfg, iq_stOut := _stOut);

// 결과 내기 (다른 경로 유닛 값은 비움: Gate가 잘못 채워도 이 경로 밖으로 새지 않게)
FOR u := 1 TO GVL_PARAM.UNIT_COUNT DO
	IF (iq_aeOpMode[u] = E_OpMode.Manual) <> bManualPath THEN
		_stOut.astUnitP[u]			:= stNone;
		_stOut.astUnitQ[u]			:= stNone;
		_stOut.abNew[u]				:= FALSE;
		_stOut.abWaitNewCmd[u]		:= FALSE;
		_stOut.aeRefuse[u]			:= E_CmdRefuse.None;
	END_IF
END_FOR
q_astUnitP		:= _stOut.astUnitP;
q_astUnitQ		:= _stOut.astUnitQ;
q_astGrpP		:= _stOut.astGrpP;
q_astGrpQ		:= _stOut.astGrpQ;
q_abNew			:= _stOut.abNew;
q_aeRefuse		:= _stOut.aeRefuse;
q_anRefuseModule:= _stOut.anRefuseModule;
q_abWaitNewCmd	:= _stOut.abWaitNewCmd;

END_FUNCTION_BLOCK

// ---- 10_Core/40_Arbitration/FB_GateAuto.TcPOU
FUNCTION_BLOCK FB_GateAuto EXTENDS FB_ModuleBase IMPLEMENTS I_Gate	// 코어 기본 Auto Gate: 그대로 통과

METHOD M_Filter
VAR_INPUT
	i_stView	: ST_GateView;
END_VAR
VAR_IN_OUT CONSTANT
	iq_astUnitP		: ARRAY[1..GVL_PARAM.UNIT_COUNT] OF ST_Pick;		// 이 경로 FB_Select 결과 (다른 경로 유닛은 비활성)
	iq_astUnitQ		: ARRAY[1..GVL_PARAM.UNIT_COUNT] OF ST_Pick;
	iq_astGrpP		: ARRAY[1..GVL_PARAM.GROUP_COUNT] OF ST_Pick;
	iq_astGrpQ		: ARRAY[1..GVL_PARAM.GROUP_COUNT] OF ST_Pick;
	iq_aeOpMode		: ARRAY[1..GVL_PARAM.UNIT_COUNT] OF E_OpMode;		// 유닛 실제 운전 모드
	iq_astUnit		: ARRAY[1..GVL_PARAM.UNIT_COUNT] OF ST_UnitState;	// 유닛 상태 (실제 출력 방향·운전 상태)
	iq_astUnitCfg	: ARRAY[1..GVL_PARAM.UNIT_COUNT] OF ST_UnitCfg;
END_VAR
VAR_IN_OUT
	iq_stOut		: ST_GateOut;		// 거른 결과 (Gate가 채움. 지난 스캔 값이 남아 있음)
END_VAR
VAR
	u	: UINT;
END_VAR
iq_stOut.astUnitP	:= iq_astUnitP;
iq_stOut.astUnitQ	:= iq_astUnitQ;
iq_stOut.astGrpP	:= iq_astGrpP;
iq_stOut.astGrpQ	:= iq_astGrpQ;
FOR u := 1 TO GVL_PARAM.UNIT_COUNT DO
	iq_stOut.abNew[u]			:= iq_astUnitP[u].bNew OR iq_astUnitQ[u].bNew;
	iq_stOut.aeRefuse[u]		:= E_CmdRefuse.None;
	iq_stOut.anRefuseModule[u]	:= 0;
	iq_stOut.abWaitNewCmd[u]	:= FALSE;
END_FOR
END_METHOD

END_FUNCTION_BLOCK

// ---- 10_Core/40_Arbitration/FB_GateManual.TcPOU
FUNCTION_BLOCK FB_GateManual EXTENDS FB_ModuleBase IMPLEMENTS I_Gate	// 코어 기본 Manual Gate (Manual 유닛만): 방향 반대 새 지령 무시(앞 값 유지), 새 지령 표시, Run 뒤 새 지령 대기
// 설정 GVL_PERSIST.g_stManualCmdSet (i_stView.stManualCmdSet). 배터리 한계는 버스 제한 모듈 (FB_SocLimit)
VAR
	_abHoldUnit		: ARRAY[1..GVL_PARAM.UNIT_COUNT] OF BOOL;			// 유닛별 값: 방향 반대로 무시해서 앞 값 유지 중
	_anHoldUnit		: ARRAY[1..GVL_PARAM.UNIT_COUNT] OF UINT;			// 무시한 지령원 (이 지령원이 끊기거나 바뀌면 유지 끝)
	_abHoldGrp		: ARRAY[1..GVL_PARAM.GROUP_COUNT] OF BOOL;
	_anHoldGrp		: ARRAY[1..GVL_PARAM.GROUP_COUNT] OF UINT;
	_abWasManual	: ARRAY[1..GVL_PARAM.UNIT_COUNT] OF BOOL;		// 지난 스캔 Manual
	_bInit			: BOOL;			// 첫 스캔: 지금 상태를 기준으로 (PMS 재기동이 운전 중 장비 출력을 바꾸지 않게)
	(* 따라가기용 중간값 *)
	_afGrpAct		: ARRAY[1..GVL_PARAM.GROUP_COUNT] OF REAL;		// 수동 그룹 몫 유닛의 실제 P 합 (그룹 지령 방향 판단)
	_afGrpBand		: ARRAY[1..GVL_PARAM.GROUP_COUNT] OF REAL;		// 이 이하는 멈춘 것으로 봄
END_VAR

METHOD M_Filter
VAR_INPUT
	i_stView	: ST_GateView;
END_VAR
VAR_IN_OUT CONSTANT
	iq_astUnitP		: ARRAY[1..GVL_PARAM.UNIT_COUNT] OF ST_Pick;		// 이 경로 FB_Select 결과 (다른 경로 유닛은 비활성)
	iq_astUnitQ		: ARRAY[1..GVL_PARAM.UNIT_COUNT] OF ST_Pick;
	iq_astGrpP		: ARRAY[1..GVL_PARAM.GROUP_COUNT] OF ST_Pick;
	iq_astGrpQ		: ARRAY[1..GVL_PARAM.GROUP_COUNT] OF ST_Pick;
	iq_aeOpMode		: ARRAY[1..GVL_PARAM.UNIT_COUNT] OF E_OpMode;		// 유닛 실제 운전 모드
	iq_astUnit		: ARRAY[1..GVL_PARAM.UNIT_COUNT] OF ST_UnitState;	// 유닛 상태 (실제 출력 방향·운전 상태)
	iq_astUnitCfg	: ARRAY[1..GVL_PARAM.UNIT_COUNT] OF ST_UnitCfg;
END_VAR
VAR_IN_OUT
	iq_stOut		: ST_GateOut;		// 거른 결과 (Gate가 채움. 지난 스캔 값이 남아 있음)
END_VAR
VAR
	u				: UINT;
	g				: UINT;
	fActualP			: REAL;
	fStopBand			: REAL;
	bNewAccepted			: BOOL;
	abGrpNew		: ARRAY[1..GVL_PARAM.GROUP_COUNT] OF BOOL;		// 그룹 P 새 지령을 받아들임 또는 그룹 Q 새 지령
	abGrpRefused	: ARRAY[1..GVL_PARAM.GROUP_COUNT] OF BOOL;
END_VAR
(* 0) 수동 그룹 몫 유닛의 실제 출력 합 (그룹 지령 방향 판단용) *)
FOR g := 1 TO GVL_PARAM.GROUP_COUNT DO
	_afGrpAct[g]		:= 0;
	_afGrpBand[g]	:= 0;
END_FOR
FOR u := 1 TO GVL_PARAM.UNIT_COUNT DO
	g := iq_astUnitCfg[u].nGroup;
	IF g >= 1 AND g <= GVL_PARAM.GROUP_COUNT AND iq_aeOpMode[u] = E_OpMode.Manual AND NOT iq_astUnitP[u].bActive THEN
		IF iq_astUnit[u].stP.bValid THEN
			_afGrpAct[g] := _afGrpAct[g] + iq_astUnit[u].stP.fValue;
		END_IF
		_afGrpBand[g] := _afGrpBand[g] + iq_astUnitCfg[u].fPRated * i_stView.stManualCmdSet.fDirBand / 100.0;
	END_IF
END_FOR

(* 1) 수동 그룹 값: 방향 반대 새 지령은 무시하고 앞 값 유지 *)
FOR g := 1 TO GVL_PARAM.GROUP_COUNT DO
	abGrpNew[g]		:= FALSE;
	abGrpRefused[g]	:= FALSE;
	IF iq_astGrpP[g].bNew THEN
		IF i_stView.stManualCmdSet.bReverse AND M_Reversed(iq_astGrpP[g], _afGrpAct[g], _afGrpBand[g]) THEN
			_abHoldGrp[g]	:= TRUE;
			_anHoldGrp[g]	:= iq_astGrpP[g].nModule;
			abGrpRefused[g]	:= TRUE;
		ELSE
			_abHoldGrp[g]	:= FALSE;
			abGrpNew[g]		:= TRUE;
		END_IF
	ELSIF NOT iq_astGrpP[g].bActive OR iq_astGrpP[g].nModule <> _anHoldGrp[g] THEN
		_abHoldGrp[g] := FALSE;
	END_IF
	IF NOT _abHoldGrp[g] THEN
		iq_stOut.astGrpP[g] := iq_astGrpP[g];
	END_IF
	iq_stOut.astGrpP[g].bNew	:= abGrpNew[g];
	iq_stOut.astGrpQ[g]			:= iq_astGrpQ[g];
	abGrpNew[g]				:= abGrpNew[g] OR iq_astGrpQ[g].bNew;
END_FOR

(* 2) 유닛별 값, 새 지령 표시, 배터리 한계 *)
FOR u := 1 TO GVL_PARAM.UNIT_COUNT DO
	g		:= iq_astUnitCfg[u].nGroup;
	fStopBand	:= iq_astUnitCfg[u].fPRated * i_stView.stManualCmdSet.fDirBand / 100.0;
	fActualP	:= 0;
	IF iq_astUnit[u].stP.bValid THEN
		fActualP := iq_astUnit[u].stP.fValue;
	END_IF

	bNewAccepted := FALSE;
	IF iq_aeOpMode[u] = E_OpMode.Manual THEN
		IF iq_astUnitP[u].bNew THEN
			IF i_stView.stManualCmdSet.bReverse AND M_Reversed(iq_astUnitP[u], fActualP, fStopBand) THEN
				_abHoldUnit[u]			:= TRUE;
				_anHoldUnit[u]			:= iq_astUnitP[u].nModule;
				iq_stOut.aeRefuse[u]			:= E_CmdRefuse.Reversed;
				iq_stOut.anRefuseModule[u]		:= iq_astUnitP[u].nModule;
			ELSE
				_abHoldUnit[u]	:= FALSE;
				bNewAccepted			:= TRUE;
			END_IF
		ELSIF NOT iq_astUnitP[u].bActive OR iq_astUnitP[u].nModule <> _anHoldUnit[u] THEN
			_abHoldUnit[u] := FALSE;
		END_IF
		bNewAccepted := bNewAccepted OR iq_astUnitQ[u].bNew;
		IF g >= 1 AND g <= GVL_PARAM.GROUP_COUNT THEN
			IF NOT iq_astUnitP[u].bActive AND abGrpRefused[g] THEN
				iq_stOut.aeRefuse[u]			:= E_CmdRefuse.Reversed;
				iq_stOut.anRefuseModule[u]		:= iq_astGrpP[g].nModule;
			END_IF
			bNewAccepted := bNewAccepted OR abGrpNew[g];
		END_IF
		IF bNewAccepted THEN
			iq_stOut.aeRefuse[u] := E_CmdRefuse.None;
		END_IF
	ELSE
		_abHoldUnit[u]	:= FALSE;
		iq_stOut.aeRefuse[u]	:= E_CmdRefuse.None;
	END_IF
	iq_stOut.abNew[u] := bNewAccepted;

	// Manual 지령은 활성(Run·대기)을 확인한 뒤 들어온 것만 씀: 활성이 아니거나 Manual로 막 들어오면 새 지령이 올 때까지 0
	// (PMS 시작 첫 스캔은 지금 상태를 기준으로만 삼음: 운전 중 장비 출력을 바꾸지 않게)
	IF NOT _bInit THEN
		_abWasManual[u] := iq_aeOpMode[u] = E_OpMode.Manual;
	END_IF
	IF i_stView.stManualCmdSet.bClearOnStop AND iq_aeOpMode[u] = E_OpMode.Manual THEN
		IF NOT (iq_astUnit[u].eRunState = E_RunState.Run OR iq_astUnit[u].eRunState = E_RunState.Standby) OR NOT _abWasManual[u] THEN
			iq_stOut.abWaitNewCmd[u] := TRUE;
		ELSIF bNewAccepted THEN
			iq_stOut.abWaitNewCmd[u] := FALSE;
		END_IF
	ELSE
		iq_stOut.abWaitNewCmd[u] := FALSE;
	END_IF
	_abWasManual[u] := iq_aeOpMode[u] = E_OpMode.Manual;

	IF NOT _abHoldUnit[u] THEN
		iq_stOut.astUnitP[u] := iq_astUnitP[u];
	END_IF
	iq_stOut.astUnitQ[u] := iq_astUnitQ[u];
END_FOR
_bInit := TRUE;
END_METHOD

METHOD PRIVATE M_Reversed : BOOL		// 새 값이 지금 출력 방향과 반대인가 (멈춰 있거나 0이면 아님)
VAR_INPUT
	i_stPick	: ST_Pick;
	i_fActualP		: REAL;			// 지금 실제 P
	i_fStopBand		: REAL;			// 이 이하는 멈춘 것으로 봄
END_VAR
M_Reversed := i_stPick.bActive AND ABS(i_fActualP) > i_fStopBand AND i_stPick.fValue * i_fActualP < 0;
END_METHOD

END_FUNCTION_BLOCK

// ---- 10_Core/40_Arbitration/FB_OutputReady.TcPOU
FUNCTION_BLOCK FB_OutputReady	// 유닛마다 지금 출력(P·Q)을 낼 수 있는지 한 번 정함. 성형(램프 기준)·분배(대상)·디스패처(Manual 쓰기 시점)는 이 결과만 씀
// 출력 가능 = 가용 + 장비 활성(Run·대기) + 정지 진행 중 아님 + 모드 전환 아님 + Manual 새 지령 대기 아님
VAR_IN_OUT CONSTANT
	iq_astAvail	: ARRAY[1..GVL_PARAM.UNIT_COUNT] OF ST_UnitAvail;	// FB_UnitAvail
	iq_astUnit	: ARRAY[1..GVL_PARAM.UNIT_COUNT] OF ST_UnitState;	// 장비 실제 상태
	iq_abStopping	: ARRAY[1..GVL_PARAM.UNIT_COUNT] OF BOOL;	// 정지 진행 중 (fbSequencer.q_abStopping, 지난 스캔)
	iq_abSwitching	: ARRAY[1..GVL_PARAM.UNIT_COUNT] OF BOOL;	// 모드 전환 중 (FB_ModeSwitch)
	iq_abManualWaitNewCmd	: ARRAY[1..GVL_PARAM.UNIT_COUNT] OF BOOL;	// Manual 새 지령 대기 (fbManualGate)
END_VAR
VAR_OUTPUT
	q_abReady	: ARRAY[1..GVL_PARAM.UNIT_COUNT] OF BOOL;	// 출력 가능
	q_aeNotReadyBy	: ARRAY[1..GVL_PARAM.UNIT_COUNT] OF E_UnitLimitBy;	// 못 내는 이유 (None = 출력 가능): NotAvail / ModeSwitch / WaitManualCmd / NotRun
END_VAR
VAR_TEMP
	u	: UINT;
END_VAR

FOR u := 1 TO GVL_PARAM.UNIT_COUNT DO
	IF NOT iq_astAvail[u].bAvail THEN
		q_aeNotReadyBy[u] := E_UnitLimitBy.NotAvail;
	ELSIF iq_abSwitching[u] THEN
		q_aeNotReadyBy[u] := E_UnitLimitBy.ModeSwitch;
	ELSIF iq_abManualWaitNewCmd[u] THEN
		q_aeNotReadyBy[u] := E_UnitLimitBy.WaitManualCmd;
	ELSIF iq_abStopping[u] OR NOT (iq_astUnit[u].eRunState = E_RunState.Run OR iq_astUnit[u].eRunState = E_RunState.Standby) THEN
		q_aeNotReadyBy[u] := E_UnitLimitBy.NotRun;
	ELSE
		q_aeNotReadyBy[u] := E_UnitLimitBy.None;
	END_IF
	q_abReady[u] := q_aeNotReadyBy[u] = E_UnitLimitBy.None;
END_FOR

END_FUNCTION_BLOCK

// ---- 10_Core/40_Arbitration/FB_LimitEval.TcPOU
FUNCTION_BLOCK FB_LimitEval		// 제한 모듈·보정 모듈을 그룹마다 한 번씩 평가 (Auto·Manual 성형이 같은 결과를 씀. 모듈 타이머가 두 번 돌지 않게)
VAR_IN_OUT CONSTANT
	iq_astView		: ARRAY[1..GVL_PARAM.GROUP_COUNT] OF ST_GroupView;
	iq_astLimitReg	: ARRAY[1..GVL_PARAM.LIMIT_COUNT] OF ST_ModuleReg;
	iq_astCompReg	: ARRAY[1..GVL_PARAM.COMP_COUNT] OF ST_ModuleReg;
END_VAR
VAR_IN_OUT
	iq_aipLimit		: ARRAY[1..GVL_PARAM.LIMIT_COUNT] OF I_LimitRule;
	iq_aipComp		: ARRAY[1..GVL_PARAM.COMP_COUNT] OF I_Compensator;
END_VAR
VAR_OUTPUT
	q_aabOn			: ARRAY[1..GVL_PARAM.GROUP_COUNT, 1..GVL_PARAM.LIMIT_COUNT] OF BOOL;		// 이 그룹에 걸린 제한 모듈
	q_aastLim		: ARRAY[1..GVL_PARAM.GROUP_COUNT, 1..GVL_PARAM.LIMIT_COUNT] OF ST_LimitOut;
	q_aaeBasis		: ARRAY[1..GVL_PARAM.GROUP_COUNT, 1..GVL_PARAM.LIMIT_COUNT] OF E_LimitBasis;
	q_aanModule		: ARRAY[1..GVL_PARAM.GROUP_COUNT, 1..GVL_PARAM.LIMIT_COUNT] OF UINT;
	q_abPccManual	: ARRAY[1..GVL_PARAM.LIMIT_COUNT] OF BOOL;		// 모듈 등록 bManual: 접속점 기준 모듈을 Manual 경로에도 적용
	q_abResume		: ARRAY[1..GVL_PARAM.GROUP_COUNT] OF BOOL;		// 재개 중인 제한 모듈 있음 (재개 램프율)
	q_afPComp		: ARRAY[1..GVL_PARAM.GROUP_COUNT] OF REAL;		// kW, 보정 합
	q_afQComp		: ARRAY[1..GVL_PARAM.GROUP_COUNT] OF REAL;		// kvar
END_VAR
VAR_TEMP
	g				: UINT;
	i				: UINT;
	stCompPQ		: ST_PQ;
END_VAR

FOR i := 1 TO GVL_PARAM.LIMIT_COUNT DO
	q_abPccManual[i] := iq_astLimitReg[i].bManual;
END_FOR
FOR g := 1 TO GVL_PARAM.GROUP_COUNT DO
	q_abResume[g] := FALSE;
	FOR i := 1 TO GVL_PARAM.LIMIT_COUNT DO
		q_aabOn[g, i] := FALSE;
		IF iq_aipLimit[i] <> 0 AND_THEN (iq_astLimitReg[i].bEnable
			AND (iq_astLimitReg[i].nGroup = 0 OR iq_astLimitReg[i].nGroup = g)) THEN
			q_aastLim[g, i]		:= iq_aipLimit[i].M_Evaluate(iq_astView[g]);
			// 제한은 줄이기만 함: 0은 항상 범위 안 (모듈이 출력을 강제하지 못함)
			q_aastLim[g, i].stP	:= F_LimitKeepZero(q_aastLim[g, i].stP);
			q_aastLim[g, i].stQ	:= F_LimitKeepZero(q_aastLim[g, i].stQ);
			q_aaeBasis[g, i]	:= iq_aipLimit[i].Basis;
			q_aanModule[g, i]	:= iq_aipLimit[i].ModuleId;
			q_aabOn[g, i]		:= TRUE;
			q_abResume[g]		:= q_abResume[g] OR q_aastLim[g, i].bResume;
		END_IF
	END_FOR

	q_afPComp[g] := 0;
	q_afQComp[g] := 0;
	FOR i := 1 TO GVL_PARAM.COMP_COUNT DO
		IF iq_aipComp[i] <> 0 AND_THEN (iq_astCompReg[i].bEnable
			AND (iq_astCompReg[i].nGroup = 0 OR iq_astCompReg[i].nGroup = g)) THEN
			stCompPQ		:= iq_aipComp[i].M_Calc(iq_astView[g]);
			// NaN·무한대 보정값은 버림 (램프 기준·Q 필터에 들어가면 풀리지 않음)
			IF F_CmdOk(stCompPQ.fP, 0) THEN q_afPComp[g] := q_afPComp[g] + stCompPQ.fP; END_IF
			IF F_CmdOk(stCompPQ.fQ, 0) THEN q_afQComp[g] := q_afQComp[g] + stCompPQ.fQ; END_IF
		END_IF
	END_FOR
END_FOR

END_FUNCTION_BLOCK

// ---- 10_Core/40_Arbitration/FB_ShapePath.TcPOU
FUNCTION_BLOCK FB_ShapePath		// 지령 다듬기, 경로 하나 (MAIN에 fbManualShape·fbAutoShape 두 개). P는 램프 → 접속점 제한 → 보정 → 설비 제한, Q는 필터 → 제한
// Auto·Manual이 같은 코드. Manual(i_bManual = TRUE)은 그룹 Manual 정책(ST_ManualPolicy)에서 켠 단계만 적용
// 유닛 지령이 기본: 그룹 지령이 없으면 이 경로 유닛 지령 합(유닛별 램프 후)을 목표로 같은 제한을 건다
// Auto는 Manual을 먼저 계산한 결과(iq_afOtherGrpP/Q)를 받아 접속점 제한을 그룹 전체로 보고, 결과에서 Manual 몫을 뺌
// 설비 제한의 정격·배터리 줄과 Q 정격은 FB_EquipmentLimits의 그룹 설비 범위 (유닛 한도 합, 버스별 배터리 한도)
VAR_INPUT
	i_bManual			: BOOL;			// TRUE = Manual 경로, FALSE = Auto 경로 (인스턴스마다 고정)
END_VAR
VAR_IN_OUT CONSTANT
	iq_astView			: ARRAY[1..GVL_PARAM.GROUP_COUNT] OF ST_GroupView;
	iq_astGroupSet		: ARRAY[1..GVL_PARAM.GROUP_COUNT] OF ST_GroupSet;
	iq_astManualPolicy	: ARRAY[1..GVL_PARAM.GROUP_COUNT] OF ST_ManualPolicy;	// Manual 경로만 씀
	iq_astUnitCfg		: ARRAY[1..GVL_PARAM.UNIT_COUNT] OF ST_UnitCfg;
	iq_aeOpMode			: ARRAY[1..GVL_PARAM.UNIT_COUNT] OF E_OpMode;			// 실제 운전 모드
	iq_abOutputReady	: ARRAY[1..GVL_PARAM.UNIT_COUNT] OF BOOL;	// 유닛 출력 가능 (FB_OutputReady). 못 내면 성형 값 0 → 기동하면 0부터 램프
	(* 이 경로 지령 (Gate 결과) *)
	iq_astUnitP			: ARRAY[1..GVL_PARAM.UNIT_COUNT] OF ST_Pick;
	iq_astUnitQ			: ARRAY[1..GVL_PARAM.UNIT_COUNT] OF ST_Pick;
	iq_astGrpP			: ARRAY[1..GVL_PARAM.GROUP_COUNT] OF ST_Pick;
	iq_astGrpQ			: ARRAY[1..GVL_PARAM.GROUP_COUNT] OF ST_Pick;
	iq_astGrpPLim		: ARRAY[1..GVL_PARAM.GROUP_COUNT] OF ST_Range;			// 이 경로 지령원 P 제한 (FB_Select)
	iq_astGrpQLim		: ARRAY[1..GVL_PARAM.GROUP_COUNT] OF ST_Range;			// 이 경로 지령원 Q 제한 (FB_Select, 접속점 기준)
	iq_afOtherGrpP		: ARRAY[1..GVL_PARAM.GROUP_COUNT] OF REAL;			// Auto: Manual 결과 (fbManualShape.q_afGrpP). Manual: 0
	iq_afOtherGrpQ		: ARRAY[1..GVL_PARAM.GROUP_COUNT] OF REAL;
	(* 제한·보정 모듈 결과 (FB_LimitEval, 그룹마다 한 번 평가) *)
	iq_aabLimOn			: ARRAY[1..GVL_PARAM.GROUP_COUNT, 1..GVL_PARAM.LIMIT_COUNT] OF BOOL;
	iq_aastLim			: ARRAY[1..GVL_PARAM.GROUP_COUNT, 1..GVL_PARAM.LIMIT_COUNT] OF ST_LimitOut;
	iq_aaeBasis			: ARRAY[1..GVL_PARAM.GROUP_COUNT, 1..GVL_PARAM.LIMIT_COUNT] OF E_LimitBasis;
	iq_aanLimModule		: ARRAY[1..GVL_PARAM.GROUP_COUNT, 1..GVL_PARAM.LIMIT_COUNT] OF UINT;
	iq_abPccManual		: ARRAY[1..GVL_PARAM.LIMIT_COUNT] OF BOOL;
	iq_abResume			: ARRAY[1..GVL_PARAM.GROUP_COUNT] OF BOOL;
	iq_afPComp			: ARRAY[1..GVL_PARAM.GROUP_COUNT] OF REAL;
	iq_afQComp	: ARRAY[1..GVL_PARAM.GROUP_COUNT] OF REAL;
	iq_astGroupEnv	: ARRAY[1..GVL_PARAM.GROUP_COUNT] OF ST_GroupEnvelope;	// 그룹 설비 범위 (FB_EquipmentLimits)
END_VAR
VAR_OUTPUT
	q_afGrpP		: ARRAY[1..GVL_PARAM.GROUP_COUNT] OF REAL;		// kW, 이 경로 유닛 몫 합 (그룹 지령 또는 유닛 지령 합, 제한 후)
	q_afGrpQ		: ARRAY[1..GVL_PARAM.GROUP_COUNT] OF REAL;		// kvar
	q_afUnitP		: ARRAY[1..GVL_PARAM.UNIT_COUNT] OF REAL;		// kW, 이 경로 유닛별 값 (램프 후, 유닛 한도는 분배에서). 지령 없으면 0
	q_afUnitQ		: ARRAY[1..GVL_PARAM.UNIT_COUNT] OF REAL;
	q_astDiag		: ARRAY[1..GVL_PARAM.GROUP_COUNT] OF ST_ShapeDiag;
	q_abGrpPCmd		: ARRAY[1..GVL_PARAM.GROUP_COUNT] OF BOOL;		// 이 경로 그룹 P 지령 있음 (제어용: 분배가 그룹 몫을 나눌지)
	q_abGrpQCmd		: ARRAY[1..GVL_PARAM.GROUP_COUNT] OF BOOL;
	q_abFollow		: ARRAY[1..GVL_PARAM.UNIT_COUNT] OF BOOL;		// 이 경로 유닛 지령을 다시 써야 함 (램프 중 또는 제한에 걸림). 디스패처는 Manual 것만 씀
END_VAR
VAR
	_afRef			: ARRAY[1..GVL_PARAM.GROUP_COUNT] OF REAL;		// 그룹 지령 램프 기준 = 지난 스캔 결과 (접속점 기준)
	_afbQFilter		: ARRAY[1..GVL_PARAM.GROUP_COUNT] OF FB_Lpf;
	(* 이번 그룹 값 (메서드에서 씀) *)
	_stEnv	: ST_GroupEnvelope;	// 이번 그룹 설비 범위
	_abLimOn		: ARRAY[1..GVL_PARAM.LIMIT_COUNT] OF BOOL;
	_astLim			: ARRAY[1..GVL_PARAM.LIMIT_COUNT] OF ST_LimitOut;
	_aeBasis		: ARRAY[1..GVL_PARAM.LIMIT_COUNT] OF E_LimitBasis;
	_anLimModule	: ARRAY[1..GVL_PARAM.LIMIT_COUNT] OF UINT;
	_abPccManual	: ARRAY[1..GVL_PARAM.LIMIT_COUNT] OF BOOL;
	_stTrace		: ST_PTrace;		// P 추적표 (메서드에서 채움)
	_astApply		: ARRAY[1..GVL_PARAM.GROUP_COUNT] OF ST_ManualPolicy;	// 그룹마다 적용할 단계 (Auto는 APPLY_ALL)
	_stApply		: ST_ManualPolicy;	// 이번 그룹 것 (메서드에서 씀)
	_stGrpP			: ST_Pick;
	_stGrpQ			: ST_Pick;
	_stSrcLim		: ST_Range;
	_stQSrcLim		: ST_Range;		// 지령원 Q 제한
	_bUnitPCmd		: BOOL;
	_fUnitPReq		: REAL;			// 유닛 P 지령 합 (램프 전)
	_fUnitPSum		: REAL;			// 유닛 P 지령 합 (램프 후)
	_bUnitQCmd		: BOOL;
	_fUnitQSum		: REAL;
	_fOtherP		: REAL;			// 접속점 제한에 같이 넣는 다른 경로 몫
	_fOtherQ		: REAL;
	_fPComp			: REAL;
	_fQComp			: REAL;
	_fUp			: REAL;			// 램프율 (재개 포함)
	_fDn			: REAL;
	_tQFilter		: TIME;
END_VAR
VAR CONSTANT
	APPLY_ALL		: ST_ManualPolicy := (bRamp := TRUE, bSrcLimit := TRUE, bPccLimit := TRUE, bComp := TRUE, bDevLimit := TRUE, bRating := TRUE, bBatLimit := TRUE);	// Auto 경로: 모든 단계 (ST_ManualPolicy에 칸을 더하면 여기도)
END_VAR
VAR_TEMP
	g				: UINT;
	u				: UINT;
	i				: UINT;
	abHasAuto		: ARRAY[1..GVL_PARAM.GROUP_COUNT] OF BOOL;		// 그룹에 Auto 유닛이 있음
	bInPath			: BOOL;
	afUp			: ARRAY[1..GVL_PARAM.GROUP_COUNT] OF REAL;		// 램프율 (램프 꺼짐이면 0)
	afDn			: ARRAY[1..GVL_PARAM.GROUP_COUNT] OF REAL;
	abGrpFollow		: ARRAY[1..GVL_PARAM.GROUP_COUNT] OF BOOL;
	abPathRun		: ARRAY[1..GVL_PARAM.GROUP_COUNT] OF BOOL;		// 그룹에 이 경로의 출력 낼 수 있는 유닛이 있음
	fShare			: REAL;
	stDiag			: ST_ShapeDiag;
END_VAR

(* 0) 그룹마다 적용할 단계와 램프율. Auto = 전부, Manual = 그룹 Manual 정책 *)
FOR g := 1 TO GVL_PARAM.GROUP_COUNT DO
	abHasAuto[g] := FALSE;
END_FOR
FOR u := 1 TO GVL_PARAM.UNIT_COUNT DO
	g := iq_astUnitCfg[u].nGroup;
	IF g >= 1 AND g <= GVL_PARAM.GROUP_COUNT AND iq_aeOpMode[u] <> E_OpMode.Manual THEN
		abHasAuto[g] := TRUE;
	END_IF
END_FOR
FOR g := 1 TO GVL_PARAM.GROUP_COUNT DO
	IF i_bManual THEN
		_astApply[g]		:= iq_astManualPolicy[g];
		_astApply[g].bComp	:= _astApply[g].bComp AND NOT abHasAuto[g];		// 같은 그룹에 Auto가 있으면 보정은 Auto 쪽에만 (두 번 더하지 않게)
	ELSE
		_astApply[g]		:= APPLY_ALL;
	END_IF
	afUp[g] := 0;
	afDn[g] := 0;
	IF iq_astGroupSet[g].bRamp AND _astApply[g].bRamp THEN		// 램프가 꺼져 있으면 램프율과 관계없이 바로 목표
		afUp[g] := iq_astGroupSet[g].fRampUp;
		afDn[g] := iq_astGroupSet[g].fRampDn;
	END_IF
END_FOR

(* 1) 유닛 지령: 램프만 (유닛 몫 램프율 = 그룹 램프율 × 유닛 정격 비율). 유닛 한도는 분배에서.
   그룹 지령이 없을 때 그룹 목표가 이 값의 합이라 먼저 계산. 램프 기준 = 지난 스캔 값.
   출력을 못 내는 유닛(멈춤·전환 중·새 지령 대기)은 0: 기동하면 0부터 램프 (계단처럼 튀지 않게) *)
FOR g := 1 TO GVL_PARAM.GROUP_COUNT DO
	abPathRun[g] := FALSE;
END_FOR
FOR u := 1 TO GVL_PARAM.UNIT_COUNT DO
	g := iq_astUnitCfg[u].nGroup;
	
	IF iq_abOutputReady[u] AND (iq_aeOpMode[u] = E_OpMode.Manual) = i_bManual AND g >= 1 AND g <= GVL_PARAM.GROUP_COUNT THEN
		abPathRun[g] := TRUE;
	END_IF
	IF iq_astUnitP[u].bActive AND iq_abOutputReady[u] AND g >= 1 AND g <= GVL_PARAM.GROUP_COUNT THEN
		fShare := 1.0;
		IF iq_astView[g].fPRatedSum > 0 THEN
			fShare := iq_astUnitCfg[u].fPRated / iq_astView[g].fPRatedSum;
		END_IF
		q_afUnitP[u] := F_RampStep(iq_astUnitP[u].fValue, q_afUnitP[u], afUp[g] * fShare, afDn[g] * fShare);
	ELSE
		q_afUnitP[u] := 0;
	END_IF
	q_afUnitQ[u] := SEL(iq_astUnitQ[u].bActive AND iq_abOutputReady[u], 0.0, iq_astUnitQ[u].fValue);	// P처럼 출력 못 내는 유닛 값은 0 (그룹 Q 합에 안 들어가게)
END_FOR

(* 2) 그룹마다: 적용할 단계, 이번 그룹 값 → M_ShapePath *)
FOR g := 1 TO GVL_PARAM.GROUP_COUNT DO
	_stEnv := iq_astGroupEnv[g];
	FOR i := 1 TO GVL_PARAM.LIMIT_COUNT DO
		_abLimOn[i]		:= iq_aabLimOn[g, i];
		_astLim[i]		:= iq_aastLim[g, i];
		_aeBasis[i]		:= iq_aaeBasis[g, i];
		_anLimModule[i]	:= iq_aanLimModule[g, i];
		_abPccManual[i]	:= iq_abPccManual[i];
	END_FOR
	_fPComp		:= iq_afPComp[g];
	_fQComp		:= iq_afQComp[g];
	_fUp		:= afUp[g];
	IF iq_astGroupSet[g].bRamp AND _astApply[g].bRamp AND (iq_abResume[g] OR iq_astGroupEnv[g].bResume) AND iq_astGroupSet[g].fRampResume > 0 THEN
		_fUp := iq_astGroupSet[g].fRampResume;
	END_IF
	_fDn		:= afDn[g];
	_tQFilter	:= iq_astGroupSet[g].tQFilter;

	_stApply	:= _astApply[g];
	// 이 경로 유닛이 하나도 출력을 못 내면 그룹 지령 램프 기준을 "이 경로 몫 0"으로 (다시 기동하면 0부터 램프)
	IF NOT abPathRun[g] THEN
		_afRef[g] := iq_afOtherGrpP[g] - SEL(_stApply.bComp, 0.0, iq_afPComp[g]);
	END_IF

	_stGrpP		:= iq_astGrpP[g];
	_stGrpQ		:= iq_astGrpQ[g];
	_stSrcLim	:= iq_astGrpPLim[g];
	_stQSrcLim	:= iq_astGrpQLim[g];
	_fOtherP	:= iq_afOtherGrpP[g];
	_fOtherQ	:= iq_afOtherGrpQ[g];
	_bUnitPCmd	:= FALSE;
	_fUnitPReq	:= 0;
	_fUnitPSum	:= 0;
	_bUnitQCmd	:= FALSE;
	_fUnitQSum	:= 0;
	FOR u := 1 TO GVL_PARAM.UNIT_COUNT DO
		IF iq_astUnitCfg[u].nGroup = g THEN
			IF iq_astUnitP[u].bActive THEN
				_bUnitPCmd	:= TRUE;
				_fUnitPReq	:= _fUnitPReq + iq_astUnitP[u].fValue;
				_fUnitPSum	:= _fUnitPSum + q_afUnitP[u];
			END_IF
			IF iq_astUnitQ[u].bActive THEN
				_bUnitQCmd	:= TRUE;
				_fUnitQSum	:= _fUnitQSum + q_afUnitQ[u];
			END_IF
		END_IF
	END_FOR

	stDiag := M_ShapePath(g);
	q_astDiag[g]	:= stDiag;
	q_abGrpPCmd[g]	:= _stGrpP.bActive;
	q_abGrpQCmd[g]	:= _stGrpQ.bActive;
	q_afGrpP[g]		:= stDiag.fPOut;
	q_afGrpQ[g]		:= stDiag.stQ.fOut - _fOtherQ;
	abGrpFollow[g]	:= ABS(stDiag.fPRamped - stDiag.fPReq) > 0.001 OR stDiag.stPcc.bClamped OR stDiag.stDev.bClamped OR stDiag.stQ.bClamped;
END_FOR

(* 3) 추종 표시: 유닛별 값 램프 중, 또는 이 경로 그룹 값이 램프 중·제한 *)
FOR u := 1 TO GVL_PARAM.UNIT_COUNT DO
	g := iq_astUnitCfg[u].nGroup;
	bInPath := (iq_aeOpMode[u] = E_OpMode.Manual) = i_bManual;
	q_abFollow[u] := iq_abOutputReady[u] AND iq_astUnitP[u].bActive AND q_afUnitP[u] <> iq_astUnitP[u].fValue;
	IF g >= 1 AND g <= GVL_PARAM.GROUP_COUNT AND bInPath AND iq_abOutputReady[u] THEN
		q_abFollow[u] := q_abFollow[u] OR abGrpFollow[g];
	END_IF
END_FOR

METHOD PRIVATE M_ShapePath : ST_ShapeDiag		// 경로 하나(Auto 또는 Manual) 성형. Auto·Manual이 같은 순서, _stApply에서 꺼진 단계만 건너뜀
// 입력: i_bManual, _stApply, _stGrpP/Q, _stSrcLim, 유닛 합(_fUnitP*·_fUnitQSum), _fOtherP/Q, _tQFilter, _fPComp/_fQComp, _fUp/_fDn, 제한 모듈 결과
VAR_INPUT
	i_nGroup	: UINT;
END_VAR
VAR
	i			: UINT;
	fUp			: REAL;
	fDn			: REAL;
	fComp		: REAL;			// 이 경로에 더하는 P 보정
	fQComp		: REAL;
	fRef		: REAL;
	fTrace		: REAL;
	tTau		: TIME;
	stRng		: ST_Range;
	stQRng		: ST_Range;
	stOne		: ST_Range;		// 모듈 하나의 범위 (추적표)
	stQLim		: ST_Limit;		// 접속점 기준 모듈 Q 제한을 설비 기준으로 옮긴 값
	stDiag		: ST_ShapeDiag;
END_VAR
fUp		:= SEL(_stApply.bRamp, 0.0, _fUp);
fDn		:= SEL(_stApply.bRamp, 0.0, _fDn);
fComp	:= SEL(_stApply.bComp, 0.0, _fPComp);
fQComp	:= SEL(_stApply.bComp, 0.0, _fQComp);
stDiag.fRampUp	:= fUp;
stDiag.fRampDn	:= fDn;
stDiag.fPComp	:= fComp;

(* P: 목표 → 램프 → 접속점 제한 → 보정 → 설비 제한
   목표 = 그룹 지령 (접속점 기준). 없으면 유닛 지령 합 (유닛별로 이미 램프함) + 다른 경로 몫 - 보정 *)
stDiag.bPGroupCmd	:= _stGrpP.bActive;
stDiag.bPUnitCmd	:= _bUnitPCmd;
stDiag.nPSource		:= _stGrpP.nModule;
fRef := _afRef[i_nGroup];
IF _stGrpP.bActive THEN
	stDiag.fPReq	:= _stGrpP.fValue;
	stDiag.fPRamped	:= F_RampStep(stDiag.fPReq, fRef, fUp, fDn);
ELSE
	stDiag.fPReq	:= _fUnitPReq + _fOtherP - fComp;
	stDiag.fPRamped	:= _fUnitPSum + _fOtherP - fComp;
END_IF

(* P 추적표: 범위를 모으면서 같은 자리에서 한 줄씩 남김 (같은 단계 안의 모듈은 등록 순서대로 하나씩 자른 값, 보기용. 출력은 모은 범위로 한 번에 자름) *)
_stTrace.nCount := 0;
M_TraceSet(E_TraceStep.Request, stDiag.fPReq, stDiag.nPSource, FALSE);
IF _stApply.bRamp THEN
	M_TraceSet(E_TraceStep.Ramp, stDiag.fPRamped, 0, ABS(stDiag.fPRamped - stDiag.fPReq) > 0.001);
END_IF

// 접속점 제한: 지령원 P 제한 + 접속점 기준 모듈 (Manual은 모듈 등록 bManual인 것만)
fTrace := stDiag.fPRamped;
stRng := F_RangeOpen();
IF _stApply.bSrcLimit THEN
	stRng := _stSrcLim;
	IF _stSrcLim.nMaxModule <> 0 OR _stSrcLim.nMinModule <> 0 THEN
		fTrace := M_TraceClamp(E_TraceStep.PccLimit, fTrace, _stSrcLim);
	END_IF
END_IF
FOR i := 1 TO GVL_PARAM.LIMIT_COUNT DO
	IF M_PccLimitOn(i) THEN
		stOne	:= F_RangeAdd(F_RangeOpen(), _astLim[i].stP, _anLimModule[i]);
		stRng	:= F_RangeAdd(stRng, _astLim[i].stP, _anLimModule[i]);
		fTrace	:= M_TraceClamp(E_TraceStep.PccLimit, fTrace, stOne);
	END_IF
END_FOR
stDiag.stPccRng	:= stRng;
stDiag.stPcc	:= F_RangeClamp(stDiag.fPRamped, stRng);

// 보정
fTrace := stDiag.stPcc.fOut + fComp;
IF _stApply.bComp THEN
	M_TraceSet(E_TraceStep.Comp, fTrace, 0, FALSE);
END_IF

// 설비 제한: 그룹 설비 범위(정격·배터리) + 설비 기준 모듈 (이번 경로에서 켠 것만)
stRng := F_RangeOpen();
IF _stApply.bRating THEN
	stRng	:= F_RangeAnd(stRng, _stEnv.stRating);
	fTrace	:= M_TraceClamp(E_TraceStep.DevRating, fTrace, _stEnv.stRating);
END_IF
IF _stApply.bBatLimit THEN
	stRng	:= F_RangeAnd(stRng, _stEnv.stBattery);
	fTrace	:= M_TraceClamp(E_TraceStep.DevBattery, fTrace, _stEnv.stBattery);
END_IF
FOR i := 1 TO GVL_PARAM.LIMIT_COUNT DO
	IF M_DevLimitOn(i) THEN
		stOne	:= F_RangeAdd(F_RangeOpen(), _astLim[i].stP, _anLimModule[i]);
		stRng	:= F_RangeAdd(stRng, _astLim[i].stP, _anLimModule[i]);
		fTrace	:= M_TraceClamp(E_TraceStep.DevLimit, fTrace, stOne);
	END_IF
END_FOR
stDiag.stDevRng	:= stRng;
stDiag.stDev	:= F_RangeClamp(stDiag.stPcc.fOut + fComp, stRng);
stDiag.fPOut	:= stDiag.stDev.fOut - _fOtherP;		// 이 경로 몫
_afRef[i_nGroup] := stDiag.stDev.fOut - fComp;		// 다음 스캔 램프 기준 (접속점 기준으로 되돌림)
stDiag.stTrace := _stTrace;

(* Q: 고르기 → 응답 필터 → 제한 (지령원 Q 제한 + 정격 + 제한 모듈 Q). 다른 경로 몫을 합쳐 제한 (Auto만) *)
stQRng := F_RangeOpen();
IF _stApply.bSrcLimit THEN
	stQRng := _stQSrcLim;		// 지령원 Q 제한 (P와 같음: Manual은 정책 bSrcLimit). 접속점 기준 → 설비 기준 (보정만큼 옮김)
	IF stQRng.nMaxModule <> 0 THEN stQRng.fMax := stQRng.fMax + fQComp; END_IF
	IF stQRng.nMinModule <> 0 THEN stQRng.fMin := stQRng.fMin + fQComp; END_IF
END_IF
IF _stApply.bRating THEN
	stQRng := F_RangeAnd(stQRng, _stEnv.stQ);
END_IF
FOR i := 1 TO GVL_PARAM.LIMIT_COUNT DO
	// Q도 P와 같은 규칙: 설비 기준 모듈은 bDevLimit, 접속점 기준 모듈은 M_PccLimitOn (Manual은 bPccLimit + 모듈 bManual)
	// Q 범위는 설비 기준(접속점 + 보정)이므로 접속점 기준 모듈 값은 보정만큼 옮겨 겹침 (P는 보정 앞 단계에서 자름)
	IF M_DevLimitOn(i) THEN
		stQRng := F_RangeAdd(stQRng, _astLim[i].stQ, _anLimModule[i]);
	ELSIF M_PccLimitOn(i) THEN
		stQLim		:= _astLim[i].stQ;
		stQLim.fMax	:= stQLim.fMax + fQComp;
		stQLim.fMin	:= stQLim.fMin + fQComp;
		stQRng := F_RangeAdd(stQRng, stQLim, _anLimModule[i]);
	END_IF
END_FOR
stDiag.stQRng		:= stQRng;
stDiag.bQGroupCmd	:= _stGrpQ.bActive;
stDiag.bQUnitCmd	:= _bUnitQCmd;
tTau := T#0S;
IF _stApply.bRamp THEN
	tTau := _tQFilter;
END_IF
// 목표 = 그룹 지령 (필터 후 + 보정). 없으면 유닛 지령 합 + 다른 경로 몫 (필터는 그 값을 따라가게만 둠)
IF _stGrpQ.bActive THEN
	_afbQFilter[i_nGroup](i_fIn := _stGrpQ.fValue, i_tTau := tTau);
	stDiag.stQ := F_RangeClamp(_afbQFilter[i_nGroup].q_fOut + fQComp, stQRng);
ELSE
	_afbQFilter[i_nGroup](i_fIn := _fUnitQSum + _fOtherQ - fQComp, i_tTau := tTau);
	stDiag.stQ := F_RangeClamp(_fUnitQSum + _fOtherQ, stQRng);
END_IF
M_ShapePath := stDiag;
END_METHOD

METHOD PRIVATE M_PccLimitOn : BOOL		// 이번 경로에 접속점 기준 모듈 i를 적용하는가
VAR_INPUT
	i_nLimit	: UINT;
END_VAR
M_PccLimitOn := _abLimOn[i_nLimit] AND _aeBasis[i_nLimit] = E_LimitBasis.Pcc
				AND (NOT i_bManual OR (_stApply.bPccLimit AND _abPccManual[i_nLimit]));
END_METHOD

METHOD PRIVATE M_DevLimitOn : BOOL		// 이번 경로에 설비 기준 모듈 i를 적용하는가 (Manual은 정책 bDevLimit)
VAR_INPUT
	i_nLimit	: UINT;
END_VAR
M_DevLimitOn := _stApply.bDevLimit AND _abLimOn[i_nLimit] AND _aeBasis[i_nLimit] = E_LimitBasis.Device;
END_METHOD

METHOD PRIVATE M_TraceSet		// 추적표에 한 줄 추가
VAR_INPUT
	i_eStep		: E_TraceStep;
	i_fValue	: REAL;
	i_nModule	: UINT;
	i_bCut		: BOOL;
END_VAR
IF _stTrace.nCount < GVL_PARAM.TRACE_STEP_MAX - 2 THEN		// 끝 두 줄(분배 후·쓴 값)은 FB_OutputDiag 몫
	_stTrace.nCount := _stTrace.nCount + 1;
	_stTrace.astStep[_stTrace.nCount].eStep		:= i_eStep;
	_stTrace.astStep[_stTrace.nCount].fValue	:= i_fValue;
	_stTrace.astStep[_stTrace.nCount].bCut		:= i_bCut;
	_stTrace.astStep[_stTrace.nCount].nModule	:= i_nModule;
	_stTrace.astStep[_stTrace.nCount].nReason	:= 0;
END_IF
END_METHOD

METHOD PRIVATE M_TraceClamp : REAL		// 범위 하나로 자르고 추적표에 한 줄. 자른 값을 돌려줌
VAR_INPUT
	i_eStep		: E_TraceStep;
	i_fIn		: REAL;
	i_stRange	: ST_Range;
END_VAR
VAR
	stClamp		: ST_Clamp;
END_VAR
stClamp := F_RangeClamp(i_fIn, i_stRange);
M_TraceSet(i_eStep, stClamp.fOut, stClamp.nModule, stClamp.bClamped);
IF _stTrace.nCount >= 1 THEN
	_stTrace.astStep[_stTrace.nCount].nReason := stClamp.nReason;
END_IF
M_TraceClamp := stClamp.fOut;
END_METHOD

END_FUNCTION_BLOCK

// ---- 10_Core/02_Util/FB_Lpf.TcPOU
FUNCTION_BLOCK FB_Lpf		// 1차 지연 필터
VAR_INPUT
	i_fIn			: REAL;
	i_tTau			: TIME;		// 시정수. T#0S면 필터 없이 통과
	i_bSync			: BOOL;		// 내부 값을 i_fSyncValue로 맞춤
	i_fSyncValue	: REAL;
END_VAR
VAR_OUTPUT
	q_fOut			: REAL;
END_VAR
VAR
	_fState			: REAL;
END_VAR
VAR_TEMP
	fDt				: REAL;		// s
	fTau			: REAL;		// s
END_VAR

fDt		:= F_CycleSec();
fTau	:= TIME_TO_REAL(i_tTau) / 1000.0;

IF i_bSync THEN
	_fState := i_fSyncValue;
ELSIF fTau <= 0 THEN
	_fState := i_fIn;
ELSE
	_fState := _fState + (fDt / (fTau + fDt)) * (i_fIn - _fState);
END_IF

q_fOut := _fState;

END_FUNCTION_BLOCK

// ---- 10_Core/02_Util/F_CycleSec.TcPOU
FUNCTION F_CycleSec : REAL		// 지금 태스크의 주기 (s)
VAR
	nTask		: DINT;
END_VAR

nTask := GETCURTASKINDEXEX();
F_CycleSec := UDINT_TO_REAL(TwinCAT_SystemInfoVarList._TaskInfo[nTask].CycleTime) * 1.0E-7;	// 100 ns 단위

END_FUNCTION

// ---- 10_Core/02_Util/F_RampStep.TcPOU
FUNCTION F_RampStep : REAL		// 기준값에서 한 스캔 동안 갈 수 있는 만큼만 목표 쪽으로
VAR_INPUT
	i_fTarget	: REAL;
	i_fRef		: REAL;			// 기준 (지난 스캔 최종 출력)
	i_fUpRate	: REAL;			// |값|이 커지는 쪽 (단위/s). 0 = 램프 없음
	i_fDnRate	: REAL;			// |값|이 작아지는 쪽 (단위/s). 0 = 램프 없음
END_VAR
VAR
	fRate		: REAL;
	fStep		: REAL;
END_VAR

IF ABS(i_fTarget) > ABS(i_fRef) AND i_fTarget * i_fRef >= 0 THEN
	fRate := i_fUpRate;
ELSE
	fRate := i_fDnRate;
END_IF

IF fRate <= 0 THEN
	F_RampStep := i_fTarget;
ELSE
	fStep		:= fRate * F_CycleSec();
	F_RampStep	:= i_fRef + LIMIT(-fStep, i_fTarget - i_fRef, fStep);
END_IF

END_FUNCTION

// ---- 10_Core/40_Arbitration/F_RangeClamp.TcPOU
FUNCTION F_RangeClamp : ST_Clamp		// 값을 범위 안으로. 상·하한이 겹치면 상한이 이김
VAR_INPUT
	i_fIn		: REAL;
	i_stRange	: ST_Range;
END_VAR

F_RangeClamp.fIn	:= i_fIn;
F_RangeClamp.fOut	:= i_fIn;
IF F_RangeClamp.fOut < i_stRange.fMin THEN
	F_RangeClamp.fOut		:= i_stRange.fMin;
	F_RangeClamp.bClamped	:= TRUE;
	F_RangeClamp.nModule	:= i_stRange.nMinModule;
	F_RangeClamp.nReason	:= i_stRange.nMinReason;
END_IF
IF F_RangeClamp.fOut > i_stRange.fMax THEN
	F_RangeClamp.fOut		:= i_stRange.fMax;
	F_RangeClamp.bClamped	:= TRUE;
	F_RangeClamp.nModule	:= i_stRange.nMaxModule;
	F_RangeClamp.nReason	:= i_stRange.nMaxReason;
END_IF

END_FUNCTION

